(* IEC 61131-3 sources: daoli-st-library/DL_Device (part 22) *)

(* ---- FB_DL_FilterSwitchLevel.st ---- *)
(*
  FB_DL_FilterSwitchLevel  —  过滤器液位/料位联锁（fail-safe LOW + 再生切换闭锁） / Filter level interlock with fail-safe LOW and regeneration interlock
  分类 Category : DL_Device
  版本 Version  : 1.0.0
  来源 Source   : t2-2-lbp — 液位联锁族零检索深化
  溯源 Origin   : clean-room 实现，未复制任何源码行
  功能 Function : 1) 传感器原始信号归一口径与 FB_DL_LevelSwitchVib 对齐（不实例化，
                  防抖上游承载）：TRUE = 介质覆盖叉体（料位高于低位）；归一取反后
                  TRUE = 低料位，防抖 tGlitch 后出 bLowLevel；
                  2) fail-safe LOW 语义：bEnable = FALSE（传感器失效/退出）→ 强制判
                  低料位（安全侧请求切换，防干转）；
                  3) 再生切换闭锁：bRegenActive 期间 + 结束后 tBlockAfter 窗内，
                  bSwReq 强制 FALSE（TOF 承载闭锁窗，闭锁沿用当拍量）；
                  4) 双表冗余可选：bRedundEn 且双表不一致持续 tDisTo → 故障级 03FE
                  独立锁存，失效安全侧强制判低。
  边界 Boundary : ① 组态闸：tGlitch/tDisTo/tBlockAfter 任一 <= 0 → 03FF 锁存；
                  ② 闭锁窗 TOF 无条件周期刷新（R7）；切换闭锁判据全当拍量；
                  ③ Device 段 0003 故障带收口：03FE/03FF 两格（分段理由见 InverterPdiPoll ②）；
                  ④ 无 GVL 依赖：纯引脚输入输出，无外部变量引用，无物理 IO 地址。
  依赖 Depends  : 与 FB_DL_LevelSwitchVib 归一口径语义对齐（不实例化）；Standard.library（TON / TOF / R_TRIG）
  码表 Error codes（Device 段 0003，窗口 041F~0421 / 故障 03FE~03FF）:
    16#0003_03FE 故障级：双表冗余失决（不一致持续 tDisTo），锁存至 bReset
    16#0003_03FF 故障级：组态非法（任一窗口域非法），锁存至 bReset
    16#0003_041F 信息级：低料位切换请求沿（bSwReq 首次 TRUE）
    16#0003_0420 信息级：再生闭锁激活（bRegenActive 期间请求被闭锁）
    16#0003_0421 信息级：冗余判定恢复正常沿（失决解除）
  修订历史 Revision :
    2026-11-19  v1.0.0  R41 首版（批次 4 · 序号 2）
*)

FUNCTION_BLOCK FB_DL_FilterSwitchLevel
VAR_INPUT
    bLvlRaw1     : BOOL := FALSE;     // 主表原始信号，TRUE = 介质覆盖叉体 [-] / Primary raw switch, TRUE = covered
    bLvlRaw2     : BOOL := TRUE;      // 备表原始信号（冗余可选），默认与主表一致口径 [-] / Secondary raw switch
    bRedundEn    : BOOL := FALSE;     // 双表冗余使能 [-] / Redundancy enable
    bRegenActive : BOOL := FALSE;     // 再生进行中 [-] / Regeneration active
    tGlitch      : TIME := T#500MS;   // 低料位确认防抖 [ms]，域 > 0 / Low-level debounce
    tDisTo       : TIME := T#2S;      // 冗余失决窗 [ms]，域 > 0 / Redundancy disagreement window
    tBlockAfter  : TIME := T#5S;      // 再生结束后闭锁延时 [ms]，域 > 0 / Post-regen interlock delay
    bEnable      : BOOL := TRUE;      // 传感器处理使能，FALSE = 失效安全侧 [-] / Sensor enable, FALSE = fail-safe
    bReset       : BOOL := FALSE;     // 复位，上升沿清故障锁存 / Reset edge clears fault latch
END_VAR
VAR_OUTPUT
    bLowLevel    : BOOL;              // 归一低料位判定（fail-safe 口径）[-] / Normalized low-level verdict
    bSwReq       : BOOL;              // 再生切换请求（闭锁窗内强制 FALSE）[-] / Switch request, forced off in interlock
    bBlock       : BOOL;              // 闭锁窗激活标志 [-] / Interlock active flag
    bError       : BOOL;              // 故障锁存标志 / Fault latch flag
    nErrId       : UDINT;             // 事件码，0 = 无事件 / Event code
END_VAR
VAR
    tonLowDeb    : TON;               // 低料位防抖定时器，无条件周期刷新 / Low-level debounce timer
    tonDisTo     : TON;               // 冗余失决定时器（专用超时命名），无条件刷新 / Disagreement timer
    tofBlock     : TOF;               // 再生闭锁窗（TOF 承载再生后延时），无条件刷新 / Post-regen interlock timer
    rtReset      : R_TRIG;            // 复位沿实例，无条件刷新 / Reset edge instance
    _bLowNorm    : BOOL;              // 归一低料位当拍量（取反口径）/ Normalized low-level flag
    _bDisagree   : BOOL;              // 双表不一致当拍量 [-] / Disagreement current-scan flag
    _bDisLat     : BOOL;              // 失决锁存位（锁存量）/ Disagreement latch bit
    _bCfgBad     : BOOL;              // 组态锁存位（锁存量）/ Config-fault latch bit
    _uFault      : UDINT;             // 故障码锁存（锁存量）/ Latched fault code
    _uInfo       : UDINT;             // 信息码，每拍重算 / Transient info code
    _bSwReqPrev  : BOOL;              // 上拍请求镜像（请求沿判据）/ Previous request mirror
    _bBlockPrev  : BOOL;              // 上拍闭锁镜像（闭锁沿判据）/ Previous block mirror
    _bDisOkPrev  : BOOL;              // 上拍一致镜像（恢复沿判据）/ Previous agreement mirror
END_VAR

(* —— 段 0：定时器与沿实例无条件周期刷新（禁置于 IF/CASE 内） —— *)
_bLowNorm := NOT bLvlRaw1;                    // 归一取反：TRUE = 低料位（当拍量）
_bDisagree := bRedundEn AND (bLvlRaw1 <> bLvlRaw2);   // 双表不一致（当拍量）
rtReset(CLK := bReset);                       // 复位沿（每拍必调）
tonLowDeb(IN := _bLowNorm AND (NOT _bDisLat), PT := tGlitch);   // 低料位防抖（每拍必调）
tonDisTo(IN := _bDisagree, PT := tDisTo);     // 失决窗（每拍必调）
tofBlock(IN := bRegenActive, PT := tBlockAfter);  // 闭锁窗（再生期间 + 再生后延时，每拍必调）

(* —— 段 1：单拍量预清零（锁存量 _uFault/_bDisLat/_bCfgBad 不入清单，禁同拍抹除） —— *)
_uInfo := 16#0000_0000;             // 信息码每拍重算
nErrId := 16#0000_0000;             // 事件码缺省无事件

(* —— 段 2：复位沿 + 组态域闸（当拍量判据） —— *)
IF rtReset.Q THEN                   // rtReset.Q = 当拍量
    _bDisLat := FALSE;              // 清失决锁存位
    _bCfgBad := FALSE;              // 清组态锁存位
    _uFault := 16#0000_0000;        // 清故障锁存码
END_IF
IF (TIME_TO_DINT(tGlitch) <= 0) OR (TIME_TO_DINT(tDisTo) <= 0) OR (TIME_TO_DINT(tBlockAfter) <= 0) THEN
    _uFault := 16#0003_03FF;        // 故障级：组态非法
    _bCfgBad := TRUE;
END_IF

(* —— 段 3：冗余失决独立锁存与恢复（R190：失决归因唯一） —— *)
IF tonDisTo.Q AND (NOT _bDisLat) THEN
    _uFault := 16#0003_03FE;        // 故障级：双表失决锁存
    _bDisLat := TRUE;
END_IF
(* 解除式逐 BOOL 标注（R240）：rtReset.Q = 当拍量；NOT _bDisagree = 当拍量；
   均不含锁存量（_bDisLat），解除边真实可达。 *)
IF rtReset.Q AND (NOT _bDisagree) AND (NOT _bCfgBad) THEN
    _bDisLat := FALSE;              // 清失决锁存位（锁存量，仅此当拍量解除沿可清）
    _uFault := 16#0000_0000;        // 清故障锁存码（锁存量，同上唯一解除路径）
END_IF
IF (NOT _bDisagree) AND _bDisOkPrev AND bRedundEn AND (NOT _bDisLat) THEN
    _uInfo := 16#0003_0421;         // 信息级：冗余判定恢复沿
END_IF

(* —— 段 4：fail-safe LOW 归一出口（失效/失决/组态坏 → 强制判低，安全侧） —— *)
IF (NOT bEnable) OR _bDisLat OR _bCfgBad THEN
    bLowLevel := TRUE;              // 安全侧强制判低（防干转，头注释②）
ELSE
    bLowLevel := tonLowDeb.Q;       // 防抖后低料位判定
END_IF

(* —— 段 5：再生切换闭锁（闭锁判据全当拍量；TOF 电平承载再生后窗） —— *)
bBlock := bRegenActive OR tofBlock.Q;   // 闭锁窗激活（再生中或再生后延时内）
bSwReq := bLowLevel AND (NOT bBlock);   // 切换请求（闭锁窗内强制 FALSE）
IF bBlock AND (NOT _bBlockPrev) THEN
    _uInfo := 16#0003_0420;         // 信息级：再生闭锁激活
END_IF
IF bSwReq AND (NOT _bSwReqPrev) THEN
    _uInfo := 16#0003_041F;         // 信息级：切换请求沿（覆盖闭锁沿，请求优先报告）
END_IF

(* —— 段 6：出口单点映射（锁存码回放，禁同拍抹除） —— *)
IF _bDisLat OR _bCfgBad THEN
    nErrId := _uFault;              // 故障锁存码回放
ELSE
    nErrId := _uInfo;               // 信息码
END_IF
bError := _bDisLat OR _bCfgBad;     // 故障标志与锁存位同源
_bSwReqPrev := bSwReq;              // 请求沿判据快照
_bBlockPrev := bBlock;              // 闭锁沿判据快照
_bDisOkPrev := NOT _bDisagree;      // 一致镜像快照

END_FUNCTION_BLOCK

(* ---- FB_DL_FlowSwitchResponseCheck.st ---- *)
(*==============================================================================
 * 组件名称 (Component)  : FB_DL_FlowSwitchResponseCheck
 * 所属子库 (Sublibrary) : DL_Device
 * 当前版本 (Version)    : 1.0.0
 * 兼容性   (Platform)   : CODESYS 3.5+ / TwinCAT 3 / 汇川 InoProShop / 施耐德 Machine Expert
 *                         仅依赖 Standard.library（TON / R_TRIG），零厂商私有库
 * 功能描述 (Function)   : 流量开关**自身响应**校核（命令-监视-判定三段式）。① 运行指令 bRunCmd
 *                         上升沿起，tRespWin 内应出现流量开关 bFlowSw 上升沿；未出现 →
 *                         eCause = eNoResponse（开关卡死 / 管路堵塞 / 接线断）；② 指令撤销后
 *                         tDropWin 内流量信号未回落 → eCause = eStuckOn（开关粘连，常闭触点焊死）。
 *                         另输出实测响应时间 tRespMeasured（供趋势与开关劣化判断）。
 * 分工声明 (Scope)      : 本件**不判干转**（干转属主为 `FB_DL_PumpDryRunGuard` /
 *                         `FB_DL_PumpDryRunProtect`），也不判流量大小与累计量；本件只判「开关
 *                         是否按命令跟上、是否按命令放开」。干转保护需要泵曲线与最小流量阈值，
 *                         语义与本件正交，禁止互相替代。
 * 接口     (Interface)  : 输入 bRunCmd 泵/阀运行指令、bFlowSw 流量开关反馈、tRespWin 响应窗、
 *                         tDropWin 回落窗、bReset 复位；输出 bSwHealthy 开关健康位、tRespMeasured
 *                         实测响应时间（ET 锁存式）、eCause 归因、eState / bError / nErrId。
 * 边界     (Boundary)   : ① 组态闸：tRespWin <= T#0S 或 tDropWin <= T#0S → 故障锁存；
 *                         ② 响应时间测量用 **TON 的 ET 锁存**（流量沿那一拍读一次 ET 并锁存，
 *                         之后不再实时读 ET——锁存后实例继续计时会把测量值篡改，R38 范式）；
 *                         ③ TON 两枚 + R_TRIG 三枚段 0 无条件周期刷新，IN 由相位派生（R228A）；
 *                         ④ 故障相迁出唯一路径 = bReset 上升沿；⑤ 零全局耦合（无 GVL / 无物理地址）。
 * 解除式   (Release)    : bReset 上升沿 ∧ 组态合法 ∧ 当拍「指令与反馈同相」（bRunCmd 与 bFlowSw
 *                         同为真或同为假，即不处于任一异常窗，全为当拍量，R240 范式）。
 *                         自证可满足（终审两式 1）：两枚 TON 的 IN 挂相位，故障相内恒假 → Q 恒假；
 *                         现场消除卡死或粘连后指令与反馈自然同相，无恒假因子。
 * 码表     (Codes)      : 16#0003_0703 故障级：流量开关响应故障总码（组态非法 / 无响应 / 粘连 /
 *                         非法相位），锁存至 bReset 上升沿，归因由 eCause 承载（R190 单件单总码）；
 *                         16#0003_0482 信息级：响应正常（本次启动已在窗内测到响应沿）。
 *                         加码反证（R90）：响应正常时 tRespMeasured 已给出数值，但「本次启动已确认
 *                         响应」与「上一轮遗留的旧响应时间」在出口上无法区分（时间量会保持），
 *                         故立一码标记本轮已确认。
 *                         码段说明：Device 的 03xx 故障子带已占满（仅余 03C5~03C9 碎片孔洞，按
 *                         实战规则 13 禁回填），故本批新开 07xx 故障子带取 16#0003_0703；
 *                         信息级用 04xx 子带取 16#0003_0482（源码实扫为空）。分段理由即此。
 * 开源溯源 (Origin)     : 道莅自研 clean-room（参考命令-监视-判定三段式与参数域，
 *                         零代码行复制；t2-2-lbp 族）
 * 修订历史 (Revision)   : 2026-11-19  v1.0.0  R45 首版（批次 4 · 序号 17）
 *==============================================================================*)

TYPE E_DL_FsrState :
(
    eIdle     := 0,     // 待机（指令撤销且反馈已回落） / Idle, command off and feedback dropped
    eRespWait := 10,    // 响应窗内等流量信号 / Waiting for flow signal inside the response window
    eRun      := 20,    // 指令在效且流量已建立 / Command on and flow established
    eDropWait := 30,    // 回落窗内等流量信号消失 / Waiting for flow signal to drop inside the drop window
    eFault    := 90     // 故障锁存相 / Fault latched phase
);
END_TYPE

TYPE E_DL_FsrCause :
(
    eNone       := 0,   // 无故障成因 / No cause
    eCfgIllegal := 1,   // 组态非法 / Illegal configuration
    eNoResponse := 2,   // 无响应（窗内无流量沿） / No response inside the window
    eStuckOn    := 3,   // 粘连（撤销后不回落） / Stuck on, no drop after release
    ePhaseBad   := 4    // 非法相位兜底 / Illegal phase fallback
);
END_TYPE

FUNCTION_BLOCK FB_DL_FlowSwitchResponseCheck
VAR_INPUT
    bRunCmd    : BOOL := FALSE;          // 泵/阀运行指令（电平） [-] / Pump or valve run command level
    bFlowSw    : BOOL := FALSE;          // 流量开关反馈 [-] / Flow switch feedback
    tRespWin   : TIME := T#3S;           // 响应窗（指令起算），域 > T#0S [ms] / Response window, domain > T#0S [ms]
    tDropWin   : TIME := T#3S;           // 回落窗（撤令起算），域 > T#0S [ms] / Drop window, domain > T#0S [ms]
    bReset     : BOOL := FALSE;          // 复位命令，上升沿清故障 [-] / Reset command, rising edge clears fault
END_VAR
VAR_OUTPUT
    bSwHealthy   : BOOL;                 // 开关健康位（无故障且不在异常窗） [-] / Switch healthy flag
    tRespMeasured: TIME;                 // 实测响应时间（ET 锁存，锁存后不随实例计时变化） [ms] / Measured response time, latched ET [ms]
    eCause       : E_DL_FsrCause;        // 故障成因出口（R190 归因唯一） / Fault cause outlet
    eState       : E_DL_FsrState;        // 状态出口，段 6 单点映射 / State outlet
    bError       : BOOL;                 // 故障锁存标志 [-] / Fault latch flag
    nErrId       : UDINT;                // 事件码，0 = 无事件 / Event code, 0 = no event
END_VAR
VAR
    _eState      : E_DL_FsrState := E_DL_FsrState.eIdle;     // 内部相位（CASE 唯一写入目标） / Internal phase
    _eCause      : E_DL_FsrCause := E_DL_FsrCause.eNone;     // 故障成因锁存（锁存量） / Latched cause
    tonResp      : TON;                  // 响应窗计时，段 0 无条件调用 / Response window timer
    tonDrop      : TON;                  // 回落窗计时，段 0 无条件调用 / Drop window timer
    rtRun        : R_TRIG;               // 指令上升沿实例，段 0 无条件调用 / Command rising edge
    rtFlow       : R_TRIG;               // 流量上升沿实例，段 0 无条件调用 / Flow rising edge
    rtReset      : R_TRIG;               // 复位沿实例，段 0 无条件调用 / Reset edge
    _tRespLatch  : TIME;                 // 响应时间锁存槽（锁存量） [ms] / Response time latch, latched
    _bRespSeen   : BOOL;                 // 本轮已测到响应沿标记（锁存量） [-] / Response-seen flag for this run
    _bCfgBad     : BOOL;                 // 组态非法当拍量 [-] / Illegal configuration
    _bSamePhase  : BOOL;                 // 指令与反馈同相当拍量 [-] / Command and feedback in the same phase
    _bFault      : BOOL;                 // 故障锁存位（锁存量） / Latched fault bit
    _uFault      : UDINT;                // 故障码锁存（锁存量） / Latched fault code
    _uInfo       : UDINT;                // 信息码，每拍重算 / Info code, recomputed each scan
END_VAR

(* —— 段 0：当拍判据派生 + 定时器与沿实例无条件周期刷新 —— *)
_bCfgBad    := (tRespWin <= T#0S) OR (tDropWin <= T#0S);                            // 组态域闸 / Configuration gate
_bSamePhase := (bRunCmd AND bFlowSw) OR ((NOT bRunCmd) AND (NOT bFlowSw));           // 指令与反馈同相 / Command and feedback in the same phase
rtRun(CLK := bRunCmd);                                                              // 指令上升沿，每拍必调（R228A） / Command rising edge
rtFlow(CLK := bFlowSw);                                                             // 流量上升沿，每拍必调 / Flow rising edge
rtReset(CLK := bReset);                                                             // 复位沿，每拍必调 / Reset edge
tonResp(IN := (_eState = E_DL_FsrState.eRespWait), PT := tRespWin);                 // 响应窗计时（IN 由相位派生） / Response window timer
tonDrop(IN := (_eState = E_DL_FsrState.eDropWait), PT := tDropWin);                 // 回落窗计时 / Drop window timer

(* —— 段 1：单拍量预清零（锁存量不入清单，R107） —— *)
_uInfo       := 16#0000_0000;      // 信息码每拍重算 / Info recomputed every scan
bSwHealthy   := FALSE;             // 健康位每拍预清 / Healthy flag preset
tRespMeasured := _tRespLatch;      // 响应时间镜像（锁存量回放，不实时读 ET） / Response time mirror from the latch
nErrId       := 16#0000_0000;      // 事件码缺省无事件 / Event code default none
bError       := FALSE;             // 故障标志每拍预清，故障分支同拍置位（R45 配对） / Flag preset

(* —— 段 2：复位沿 + 组态域闸 —— *)
IF rtReset.Q THEN                                                        // 当拍复位沿 / current-scan reset edge
    _bFault := FALSE;                                                    // 清故障锁存位（锁存量） / Clear fault latch
    _uFault := 16#0000_0000;                                             // 清故障锁存码（锁存量） / Clear latched code
    _eCause := E_DL_FsrCause.eNone;                                      // 清成因（锁存量） / Clear latched cause
    IF _eState = E_DL_FsrState.eFault THEN
        _eState := E_DL_FsrState.eIdle;                                  // 故障相迁出唯一路径 / Sole exit from fault phase
    END_IF
END_IF
IF _bCfgBad THEN                                                         // 组态域闸 / Configuration gate
    _uFault := 16#0003_0703;                                             // 故障级：流量开关响应故障总码 / Fault-level: flow-switch fault code
    _bFault := TRUE;
    bError  := TRUE;                                                     // 故障标志同拍置位（R45 配对） / Error flag set same scan
    _eCause := E_DL_FsrCause.eCfgIllegal;                                // 归因：组态非法 / Cause: illegal configuration
END_IF

(* —— 段 3：响应时间测量（ET 只在流量沿那一拍读一次并锁存，R38 范式） —— *)
IF (NOT _bFault) AND (_eState = E_DL_FsrState.eRespWait) AND rtFlow.Q THEN
    _tRespLatch := tonResp.ET;                                           // 锁存响应时间（此后不再实时读 ET） / Latch ET once, never re-read live
    _bRespSeen := TRUE;                                                  // 本轮已确认响应 / Response confirmed for this run
    _uInfo := 16#0003_0482;                                              // 信息级：响应正常 / Info: response OK
END_IF

(* —— 段 4：无响应 / 粘连双判据（各用独立实例与独立归因，R190） —— *)
IF (NOT _bFault) AND tonResp.Q THEN                                      // 响应窗内无流量沿 → 无响应 / No flow edge inside the window
    _uFault := 16#0003_0703;
    _bFault := TRUE;
    bError  := TRUE;
    _eCause := E_DL_FsrCause.eNoResponse;                                // 归因：无响应 / Cause: no response
END_IF
IF (NOT _bFault) AND tonDrop.Q THEN                                      // 回落窗内流量未消失 → 粘连 / Flow did not drop inside the window
    _uFault := 16#0003_0703;
    _bFault := TRUE;
    bError  := TRUE;
    _eCause := E_DL_FsrCause.eStuckOn;                                   // 归因：粘连 / Cause: stuck on
END_IF

(* —— 段 5：故障解除式（R240 全当拍量） —— *)
IF rtReset.Q AND (NOT _bCfgBad) AND _bSamePhase THEN
    _bFault := FALSE;                                                    // 清故障锁存位（锁存量） / Clear fault latch
    _uFault := 16#0000_0000;                                             // 清故障锁存码（锁存量） / Clear latched code
    _eCause := E_DL_FsrCause.eNone;                                      // 清成因（锁存量） / Clear latched cause
END_IF

(* —— 段 5A：故障锁存相位迁移闸 —— *)
IF _bFault AND (_eState <> E_DL_FsrState.eFault) THEN
    _eState := E_DL_FsrState.eFault;                                     // 锁存即入故障相 / Latch enters fault phase
END_IF

(* —— 段 6：相位机（ENUM 全成员显式标签 + ELSE 兜底，R128） —— *)
CASE _eState OF

E_DL_FsrState.eIdle:
    IF rtRun.Q AND (NOT _bFault) THEN                                    // 出口 1：收到运行指令 / Run command received
        _bRespSeen := FALSE;                                             // 新一轮响应测量重新武装 / Re-arm response measurement
        _eState := E_DL_FsrState.eRespWait;
    ELSIF bFlowSw AND (NOT bRunCmd) THEN                                 // 出口 2：无令而流量已在（越序，交由回落链监视） / Flow on without command
        _eState := E_DL_FsrState.eDropWait;
    ELSIF _bFault THEN                                                   // 出口 3：故障锁存 / Fault latched
        _eState := E_DL_FsrState.eFault;
    END_IF

E_DL_FsrState.eRespWait:
    IF rtFlow.Q THEN                                                     // 出口 1：窗内出现流量沿 / Flow edge inside the window
        _eState := E_DL_FsrState.eRun;
    ELSIF NOT bRunCmd THEN                                               // 出口 2：指令撤销（前置消失，R98） / Command released
        _eState := E_DL_FsrState.eIdle;
    END_IF

E_DL_FsrState.eRun:
    IF NOT bRunCmd THEN                                                  // 出口 1：撤销指令，进回落窗 / Command released, enter drop window
        _eState := E_DL_FsrState.eDropWait;
    ELSIF NOT bFlowSw THEN                                               // 出口 2：运行中流量消失（前置消失，R98） / Flow lost while running
        _eState := E_DL_FsrState.eRespWait;
    END_IF

E_DL_FsrState.eDropWait:
    IF NOT bFlowSw THEN                                                  // 出口 1：流量已回落 / Flow dropped
        _eState := E_DL_FsrState.eIdle;
    ELSIF bRunCmd THEN                                                   // 出口 2：指令重新来（前置消失，R98） / Command came back
        _eState := E_DL_FsrState.eRespWait;
    END_IF

E_DL_FsrState.eFault:
    ;                                                                     // 故障相：仅段 5 复位沿可迁出 / Only the reset edge leaves this phase

ELSE
    _uFault := 16#0003_0703;                                             // 故障级：非法相位兜底（归并总码） / Illegal-phase fallback
    _bFault := TRUE;
    bError  := TRUE;
    _eCause := E_DL_FsrCause.ePhaseBad;                                  // 归因：非法相位 / Cause: illegal phase
    _eState := E_DL_FsrState.eFault;

END_CASE

(* —— 段 7：出口单点映射（名实同源；锁存码回放） —— *)
bSwHealthy := (NOT _bFault) AND _bSamePhase AND _bRespSeen;              // 健康 = 无故障 ∧ 同相 ∧ 本轮已确认响应 / Healthy verdict
IF _bFault THEN
    nErrId := _uFault;                                                   // 故障锁存码回放 / Replay latched fault code
ELSE
    nErrId := _uInfo;                                                    // 信息码 / Info code
END_IF
bError := _bFault;                                                       // 故障标志与锁存同源（名实双出口，R191） / Flag from latch
eState := _eState;                                                       // 状态出口 / State outlet
eCause := _eCause;                                                       // 成因出口 / Cause outlet

END_FUNCTION_BLOCK

(* ---- FB_DL_FoupDoorSeq.st ---- *)
// =====================================================================
// FB_DL_FoupDoorSeq.st
// FOUP 开合门与载具联锁顺控（解锁-开门-载具在位-再锁定确认窗）
// FOUP door interlock sequencing with relock confirm window
// 所属子库: DL_Device    版本: v1.0.0    兼容: CODESYS V3.5+ / TwinCAT 3 / 汇川 InoProShop
// 码位: 16#0003_03DE ~ 16#0003_03E2 (本件独占 5 槽, 勿复用)
// 溯源: 道莅 clean-room 防御性实现
//       来源组标签: semiconductor, door-interlock, sequencing, foup
// 枚举属主: E_DL_FoupDoorState —— 本文件为全库唯一属主, 其他件只引用不重声明
// 修改记录: R30 初版 (ROUND_PLAN_R30 序 2)
// =====================================================================
// ---------------------------------------------------------------------
// 枚举定义: E_DL_FoupDoorState (全库唯一属主, 其他件只引用不重声明)
// ---------------------------------------------------------------------
TYPE E_DL_FoupDoorState :
(
    eIdle,          // 空闲（门锁闭等待）/ Idle, locked
    eUnlocking,     // 解锁保持中 / Unlocking
    eDoorOpen,      // 门已开等待传输 / Door open
    eTransfer,      // 载具传输中 / Transfer in progress
    eRelocking,     // 再锁定确认窗 / Relocking confirm window
    eFault          // 故障锁存 / Fault latched
);
END_TYPE

FUNCTION_BLOCK FB_DL_FoupDoorSeq
VAR_INPUT
    bEnable         : BOOL  := FALSE;   // 使能 / Enable
    bDoorClosed     : BOOL  := FALSE;   // 门磁关到位反馈 / Door closed feedback
    bDoorOpen       : BOOL  := FALSE;   // 门磁开到位反馈 / Door open feedback
    bCarrierPresent : BOOL  := FALSE;   // 载具在位检测 / Carrier present detection
    bUnlockCmd      : BOOL  := FALSE;   // 解锁命令 / Unlock command
    bLockCmd        : BOOL  := FALSE;   // 锁定命令 / Lock command
    bVacuumOk       : BOOL  := FALSE;   // 真空解锁条件就绪 / Vacuum release ready
    tUnlockHold     : TIME  := T#3S;    // 解锁保持超时窗 T#100MS~T#60S / Unlock hold timeout window [s]
    tRelockWin      : TIME  := T#5S;    // 再锁定确认窗 T#100MS~T#60S / Relock confirm window [s]
    bReset          : BOOL  := FALSE;   // 故障复位命令 / Fault reset command
END_VAR
VAR_OUTPUT
    bUnlockOut      : BOOL := FALSE;    // 解锁输出, 安全侧为假 / Unlock output, safe side FALSE
    bLockOut        : BOOL := FALSE;    // 锁定输出 / Lock output
    eState          : E_DL_FoupDoorState := E_DL_FoupDoorState.eIdle;  // 顺控状态 / Sequence state
    bTransferPermit : BOOL := FALSE;    // 载具传输允许 / Transfer permit
    eErr            : UDINT := 16#0003_03DE;  // 错误码 / Error code
END_VAR
VAR
    eErrLatch       : UDINT := 16#0003_03DE;  // 故障锁存码回放 / Latched fault code replay
    bDoorConflict   : BOOL := FALSE;    // 门磁双反馈矛盾 / Door feedback conflict
    rtrReset        : R_TRIG;           // 复位上升沿检测, 每拍无条件刷新 / Reset edge, refreshed every cycle
    tonUnlock       : TON;              // 解锁保持超时定时器, 每拍无条件刷新 / Unlock hold timer, refreshed every cycle
    tonRelock       : TON;              // 再锁定确认窗定时器, 每拍无条件刷新 / Relock window timer, refreshed every cycle
END_VAR

// ---------------------------------------------------------------------
// 代码位表（本件独占, 勿复用）:
//   16#0003_03DE 信息 顺控正常（空闲或顺控执行中）
//   16#0003_03DF 故障 解锁保持超时（解锁输出有效而门未开超时）, 解除式 = bReset 上升沿 且 门磁回到关到位 且 无矛盾反馈
//   16#0003_03E0 故障 再锁定确认窗超时（窗内门磁未回关到位）, 解除式同 03DF
//   16#0003_03E1 故障 门磁双反馈矛盾（关到位与开到位同时有效）, 解除式同 03DF
//   16#0003_03E2 故障 非法状态兜底（状态机 ELSE 拦截）, 解除式同 03DF
// ---------------------------------------------------------------------

// ---- 门磁矛盾判（最高优先级拦截）/ Door feedback conflict: highest priority ----
bDoorConflict := bDoorClosed AND bDoorOpen;     // 双反馈同有效 = 组态或接线矛盾 / Both active = conflict
IF bDoorConflict THEN
    eState    := E_DL_FoupDoorState.eFault;     // 任意相直接落故障 / Fall to fault from any phase
    eErrLatch := 16#0003_03E1;                  // 锁存矛盾码 / Latch conflict code
END_IF

// ---- 非故障相下使能撤销 → 回空闲（安全侧）/ Disable in non-fault phase returns to idle ----
IF (NOT bEnable) AND (eState <> E_DL_FoupDoorState.eFault) THEN
    eState := E_DL_FoupDoorState.eIdle;         // 退回空闲 / Return to idle
END_IF

// ---- 定时器与边沿实例无条件周期刷新（调用本身不进任何 IF 分支）/ Unconditional timer and edge refresh ----
tonUnlock(IN := (eState = E_DL_FoupDoorState.eUnlocking) AND (NOT bDoorOpen),
          PT := tUnlockHold);                   // 解锁保持计时 / Unlock hold timing
tonRelock(IN := (eState = E_DL_FoupDoorState.eRelocking) AND (NOT bDoorClosed),
          PT := tRelockWin);                    // 再锁定确认窗计时 / Relock window timing
rtrReset(CLK := bReset);                        // 复位沿检测 / Reset edge detection

// ---- 默认输出（安全侧全 0, 各相按需覆盖）/ Default outputs (safe side) ----
bUnlockOut      := FALSE;   // 解锁输出缺省断开 / Unlock default off
bLockOut        := FALSE;   // 锁定输出缺省断开 / Lock default off
bTransferPermit := FALSE;   // 传输允许缺省禁止 / Permit default denied

// ---- 状态机 / State machine ----
IF eState = E_DL_FoupDoorState.eFault THEN
    // 故障相: 输出全 0, 锁存码回放 / Fault phase: outputs all off, latch replay
    eErr := eErrLatch;
    // 解除式: bReset 上升沿 且 门磁回到关到位 且 无矛盾反馈 / Release: reset edge AND closed AND no conflict
    IF rtrReset.Q AND bDoorClosed AND (NOT bDoorOpen) AND (NOT bDoorConflict) THEN
        eState    := E_DL_FoupDoorState.eIdle;  // 解除故障回空闲 / Release to idle
        eErrLatch := 16#0003_03DE;              // 清锁存码 / Clear latch code
    END_IF
ELSE
    CASE eState OF
        E_DL_FoupDoorState.eIdle:       // 空闲: 门锁闭等待解锁命令 / Idle: locked, wait unlock
            bLockOut := bDoorClosed;    // 锁定输出随关到位反馈 / Lock output follows closed feedback
            IF bUnlockCmd AND bVacuumOk AND (NOT bDoorConflict) THEN
                eState := E_DL_FoupDoorState.eUnlocking;    // 拍 N 进入解锁相 / Enter unlocking
            END_IF
        E_DL_FoupDoorState.eUnlocking:  // 解锁保持: 输出有效等待门开 / Unlocking: output on, wait door open
            bUnlockOut := TRUE;         // 解锁输出有效 / Unlock output on
            // 本拍行为: 门开转开门相, 真空条件丢失回空闲, 超时落故障 / Open to door phase, vacuum loss to idle, timeout to fault
            IF bDoorOpen AND (NOT bDoorConflict) THEN
                eState := E_DL_FoupDoorState.eDoorOpen;     // 拍 N+1 转开门相 / To door-open phase
            ELSIF NOT bVacuumOk THEN
                eState := E_DL_FoupDoorState.eIdle;         // 真空条件丢失中止解锁 / Vacuum lost, abort unlock
            ELSIF tonUnlock.Q THEN
                eState    := E_DL_FoupDoorState.eFault;     // 解锁有效但门未开超时 / Unlock valid but not open in time
                eErrLatch := 16#0003_03DF;                  // 锁存超时码 / Latch timeout code
            END_IF
        E_DL_FoupDoorState.eDoorOpen:   // 门已开: 允许传输, 等载具在位或锁定命令 / Door open: permit, wait carrier or lock cmd
            bUnlockOut      := TRUE;    // 开门期间保持解锁 / Hold unlock while open
            bTransferPermit := TRUE;    // 允许载具传输 / Permit transfer
            IF bCarrierPresent THEN
                eState := E_DL_FoupDoorState.eTransfer;     // 载具在位转传输相 / Carrier present, to transfer
            ELSIF bLockCmd AND (NOT bDoorConflict) THEN
                eState := E_DL_FoupDoorState.eRelocking;    // 直接收到锁定命令转确认窗 / Lock cmd, to relocking
            END_IF
        E_DL_FoupDoorState.eTransfer:   // 载具传输中: 保持允许, 等锁定命令 / Transfer: permit held, wait lock cmd
            bUnlockOut      := TRUE;    // 传输期间保持解锁 / Hold unlock during transfer
            bTransferPermit := TRUE;    // 保持传输允许 / Hold transfer permit
            IF bLockCmd AND (NOT bDoorConflict) THEN
                eState := E_DL_FoupDoorState.eRelocking;    // 收到锁定命令转确认窗 / Lock cmd, to relocking
            END_IF
        E_DL_FoupDoorState.eRelocking:  // 再锁定确认窗: 门磁必须回关到位 / Relocking: door must return closed
            bLockOut := TRUE;           // 锁定输出有效 / Lock output on
            // 本拍行为: 门关到位转空闲, 窗超时落故障 / Closed to idle, window timeout to fault
            IF bDoorClosed AND (NOT bDoorConflict) THEN
                eState := E_DL_FoupDoorState.eIdle;     // 再锁定完成回空闲 / Relock done, to idle
            ELSIF tonRelock.Q THEN
                eState    := E_DL_FoupDoorState.eFault; // 确认窗内门磁未回关到位 / Door not closed in window
                eErrLatch := 16#0003_03E0;              // 锁存确认窗超时码 / Latch window timeout code
            END_IF
        ELSE                                    // 非法状态兜底拦截 / Illegal state fallback
            eState    := E_DL_FoupDoorState.eFault;     // 落故障相 / Fall to fault
            eErrLatch := 16#0003_03E2;                  // 锁存兜底码 / Latch fallback code
        END_CASE
    // 本拍错误码: 刚落故障则回放锁存码, 否则正常码 / Error code of this cycle
    IF eState = E_DL_FoupDoorState.eFault THEN
        eErr := eErrLatch;          // 回放锁存码 / Replay latch code
    ELSE
        eErr := 16#0003_03DE;       // 顺控正常 / Sequence normal
    END_IF
END_IF

END_FUNCTION_BLOCK

(* ---- FB_DL_FoupPurgeN2Flow.st ---- *)
(*
  FB_DL_FoupPurgeN2Flow  —  FOUP 氮气吹扫流量与露点监视（建立窗口 / 分级露点告警 / 注入脉冲流量计）/ FOUP N2 purge flow and dew-point supervision
  分类 Category : DL_Device
  码位 Code     : 16#03_2_0F
  版本 Version  : 1.0.0
  来源 Source   : t2-1-lgf-measurement — IEC 61131-3 标准语义的道莅防御性实现
  溯源 Origin   : LGF 测量类文档公开语义借鉴（流量带判据、露点分级），clean-room 实现，未复制源码行
  功能 Function : 1) 注入 FB_DL_PulseFlowMeter 实例（VAR_IN_OUT，只读其流量/总量/故障输出，**本件不调用其实例体**），
                     取瞬时流量与 K 系数参与判据；
                  2) 吹扫起始（bPurgeStart 上升沿）后在 tPurgeEstablish 内流量须进入 fFlowSetLpm ± fFlowTolPct% 带，
                     否则置 bEstablishTimeout（故障级 021F）；
                  3) 露点按两级判据告警：越 fDewPointMaxC 为「越限」（023F），越 fDewSevereC 为「严重越限」（024F），
                     两码独立、独立出口（R190 归因唯一）；
                  4) 露点信号质量坏或缺失时**不当作合格**：置 022F 且 bPurgeOk := FALSE（安全侧，绝不静默放行）。
  边界 Boundary : ① fFlowSetLpm <= 0 判组态错 020F（偏差百分比的分母，R45 防除零）；
                     注入流量计 fKFactor = 0 判组态错 020F 且不投运（K 系数未标定，流量读数无物理意义）；
                     露点两级门限倒置（fDewSevereC <= fDewPointMaxC）同判组态错；
                  ② 偏差百分比对 ABS 结果限幅 DL_DEV_CLAMP_PCT，防极端读数导致 REAL 溢出与 HMI 显示异常；
                  ③ bPurgeOk 的成立条件 = 建立成功 AND 流量在带 AND 露点未越限 AND 露点信号有效 AND 无故障；
                  ④ 解除式自证：_bFault 清除 = rtReset.Q（引脚可满足）；021F 另可由「流量重新入带且持续
                     tEstablishRetry」按码专清（R188 可达清除边）；023F/024F 可由露点回落按码专清；
                  ⑤ bDewPointAlarm / bDewSevereAlarm 为保持型告警位（不随单拍读数抖动），只由复位沿或回落清除。
  依赖 Depends  : FB_DL_PulseFlowMeter（DL_Device 既有件，×1 以 VAR_IN_OUT 注入）；
                  仅 Standard.library（TON / R_TRIG / ABS / MIN / MAX）
  同拍双窗配比  : tPurgeEstablish（建立窗口）与 tDewDb（露点去抖窗）不同源；配比约束
                  tDewDb <= tPurgeEstablish，保证建立窗口内露点结论至少更新一次（R100）

  码表 Error codes（本件格 03_2_0F，子码步进 +0x10）:
    16#0003_020F 故障级：组态非法（流量设定 <= 0 / K 系数 = 0 / 容差 <= 0 / 露点门限倒置 / 时间参数 <= 0）
    16#0003_021F 故障级：吹扫建立超时（tPurgeEstablish 内流量未进入容许带）
    16#0003_022F 故障级：露点信号无效（质量坏或缺失，不当作合格）
    16#0003_023F 故障级：露点越限（超 fDewPointMaxC）
    16#0003_024F 故障级：露点严重越限（超 fDewSevereC）
    16#0003_025F 故障级：状态机落 ELSE 兜底（非法相位 ID）
    16#0003_010F 信息级：吹扫建立成功，流量已入带（不置 bError）
    16#0003_011F 信息级：流量偏差瞬时越带但未超建立窗口（不置 bError）

  修订历史 Revision :
    2026-11-18  v1.0.0  R37 首版
*)

TYPE E_DL_N2PurgeState :
(
    eIdle      := 0,   // 空闲：未吹扫 / Idle, purge not started
    eEstablish := 10,  // 建立中：等流量进入容许带 / Establishing, waiting for the flow band
    ePurged    := 20,  // 吹扫中：流量与露点均在限内 / Purging, flow and dew point inside the limits
    eTimeout   := 30,  // 超时：建立窗口耗尽，等待复位 / Timed out, waiting for a reset
    eFault     := 90   // 故障：组态或信号故障锁定 / Fault, a latched configuration or signal fault
);
END_TYPE

FUNCTION_BLOCK FB_DL_FoupPurgeN2Flow
VAR_INPUT
    bEnable        : BOOL := FALSE;             // 总使能，FALSE 时 bPurgeOk 恒假 / Master enable, low level forces bPurgeOk FALSE
    bReset         : BOOL := FALSE;             // 复位，上升沿清故障与告警锁存 / Reset, clears the fault and alarm latches
    bPurgeStart    : BOOL := FALSE;             // 吹扫起始触发（上升沿受理）/ Purge start trigger, rising edge
    fFlowSetLpm    : REAL := 20.0;              // 吹扫流量设定 [L/min]，域 > 0 / Purge flow setpoint [L/min]
    fFlowTolPct    : REAL := 10.0;              // 流量容许带 [%]，域 > 0 / Flow tolerance band [%]
    fDewPointMaxC  : REAL := -40.0;             // 露点越限门限 [°C]，域 < fDewSevereC / Dew point limit [degC]
    fDewSevereC    : REAL := -20.0;             // 露点严重越限门限 [°C]，须 > fDewPointMaxC / Severe dew point limit [degC]
    fDewPointC     : REAL := -60.0;             // 露点实测值 [°C] / Measured dew point [degC]
    bDewQualityOk  : BOOL := TRUE;              // 露点信号质量（FALSE = 坏或缺失）/ Dew point signal quality, FALSE means bad
    tPurgeEstablish : TIME := T#10S;            // 吹扫建立窗口 [ms]，域 > 0 / Purge establishment window [ms]
    tEstablishRetry : TIME := T#30S;            // 入带持续窗（021F 按码专清用）[ms]，域 > 0 / In-band dwell for the code-specific clear
    tDewDb         : TIME := T#2S;              // 露点告警去抖窗 [ms]，域 > 0 / Dew point debounce [ms]
END_VAR
VAR_OUTPUT
    bPurgeOk       : BOOL;                      // 吹扫合格（建立成功且流量/露点均在限内）/ Purge acceptable
    bEstablishTimeout : BOOL;                   // 建立超时（保持型）/ Establishment timeout, held
    bDewPointAlarm : BOOL;                      // 露点越限告警（保持型）/ Dew point alarm, held
    bDewSevereAlarm : BOOL;                     // 露点严重越限告警（保持型）/ Severe dew point alarm, held
    fFlowDeviationPct : REAL;                   // 流量偏差 [%]，已限幅 / Flow deviation [%], clamped
    fFlowActualLpm : REAL;                      // 实测流量 [L/min] / Measured flow [L/min]
    bValid         : BOOL;                      // 判据可用标志 / Criteria usable
    bError         : BOOL;                      // 故障标志，派生自锁存 / Fault flag derived from the latch
    nErrId         : UDINT;                     // 事件码，0 = 无事件 / Event code, 0 = no event
    eStateOut      : E_DL_N2PurgeState;         // 状态出口，段尾单点映射 / State outlet, mapped at the tail
END_VAR
VAR_IN_OUT
    fbFlowMeter : FB_DL_PulseFlowMeter;         // 注入的脉冲流量计实例（只读输出，本件不调用其实例体）/ Injected pulse flow meter, read only
END_VAR
VAR
    tonEstablish : TON;                         // 建立窗口计时，每拍无条件调用 / Establishment window, called unconditionally
    tonInBand    : TON;                         // 入带持续计时，每拍无条件调用 / In-band dwell timer, called unconditionally
    tonDew       : TON;                         // 露点去抖计时，每拍无条件调用 / Dew point debounce, called unconditionally
    tonHeart     : TON;                         // 周期心跳窗，自复位 / Periodic heartbeat window, self-resetting
    rtReset      : R_TRIG;                      // 复位上升沿 / Reset rising edge
    rtStart      : R_TRIG;                      // 吹扫起始上升沿 / Purge start rising edge
    _eState      : E_DL_N2PurgeState := E_DL_N2PurgeState.eIdle;  // 内部相位（CASE 唯一写入目标）/ Internal phase
    _uFault      : UDINT;                       // 故障码锁存 / Latched fault code
    _uInfo       : UDINT;                       // 信息码，每拍重算 / Information code, recomputed per scan
    _bFault      : BOOL;                        // 故障锁存位 / Latched fault bit
    _bCfgBad     : BOOL;                        // 组态非法聚合 / Configuration invalid aggregate
    _bInBand     : BOOL;                        // 流量在容许带 / Flow inside the tolerance band
    _bEstTimeout : BOOL;                        // 建立超时保持量 / Held establishment-timeout value
    _bDewAlarm   : BOOL;                        // 露点越限保持量 / Held dew point alarm
    _bDewSevere  : BOOL;                        // 露点严重越限保持量 / Held severe dew point alarm
    _bDewBad     : BOOL;                        // 露点信号无效 / Dew point signal unusable
    _bEstBreak   : BOOL := TRUE;                // 建立窗口断输入一拍 / One-scan establishment break
    _bInBandBrk  : BOOL := TRUE;                // 入带计时断输入一拍 / One-scan in-band break
    _bDewBrk     : BOOL := TRUE;                // 露点去抖断输入一拍 / One-scan dew break
    _bHeartBrk   : BOOL := TRUE;                // 心跳窗断输入一拍 / One-scan heartbeat break
    _fDevRaw     : REAL;                        // 未限幅偏差 [%] / Unclamped deviation [%]
    _fKFactor    : REAL;                        // 注入流量计 K 系数 [pulses/L] / Injected K-factor [pulses/L]
END_VAR
VAR CONSTANT
    DL_DEV_CLAMP_PCT : REAL := 1000.0;   // 偏差绝对值限幅 [%] / Deviation magnitude clamp [%]
    DL_DEW_LIM_C     : REAL := 200.0;    // 露点有限性上限 [°C] / Dew point magnitude ceiling [degC]
    DL_FLOW_LIM_LPM  : REAL := 100000.0; // 流量有限性上限 [L/min] / Flow magnitude ceiling [L/min]
    DL_HEART_WINDOW  : TIME := T#2S;     // 心跳观察窗 [ms]，自复位节拍 / Heartbeat window, self-resetting
END_VAR

(* —— 段 0：定时器与边缘检测无条件周期刷新（R182：调用语句不得置于 IF / CASE 内） —— *)
rtReset(CLK := bReset);                                          // 复位上升沿，每拍必调
rtStart(CLK := bPurgeStart);                                     // 吹扫起始上升沿，每拍必调
tonHeart(IN := (NOT tonHeart.Q) AND (NOT _bHeartBrk), PT := DL_HEART_WINDOW);  // 心跳窗自复位
_bHeartBrk := FALSE;                                             // 断输入拍在调用后自清
tonEstablish(IN := (_eState = E_DL_N2PurgeState.eEstablish) AND (NOT _bEstBreak), PT := tPurgeEstablish);  // 建立窗口
_bEstBreak := FALSE;                                             // 断输入拍在调用后自清
tonInBand(IN := _bInBand AND (NOT _bInBandBrk), PT := tEstablishRetry);   // 入带持续（表达式入参）
_bInBandBrk := FALSE;                                            // 断输入拍在调用后自清
tonDew(IN := _bDewBad AND (NOT _bDewBrk), PT := tDewDb);          // 露点信号无效去抖（表达式入参）
_bDewBrk := FALSE;                                               // 断输入拍在调用后自清

(* —— 段 1：单拍量预清零（告警保持量 / 锁存不入清单，R187①） —— *)
_uInfo      := 16#0000_0000;   // 信息码每拍重算
bError      := FALSE;          // 故障出口每拍重算，段 6 由锁存派生
bValid      := FALSE;          // 可用标志缺省 FALSE
bPurgeOk    := FALSE;          // 合格出口缺省 FALSE（安全侧）
_bCfgBad    := FALSE;          // 组态非法预清零
_bInBand    := FALSE;          // 在带判据预清零
_bDewBad    := FALSE;          // 露点信号无效预清零

(* —— 段 2：复位沿清锁存与告警保持量（R188 双路径） —— *)
IF rtReset.Q THEN
    _bFault     := FALSE;            // 复位沿清锁存位
    _uFault     := 16#0000_0000;     // 复位沿清锁存码
    _bEstTimeout := FALSE;           // 清建立超时保持量
    _bDewAlarm  := FALSE;            // 清露点越限告警
    _bDewSevere := FALSE;            // 清露点严重越限告警
END_IF
IF (_uFault = 16#0003_023F) AND (NOT _bDewAlarm) THEN
    _uFault := 16#0000_0000;         // 按码专清：露点回落至越限门限以下
    _bFault := FALSE;                // 锁存位同步清
END_IF
IF (_uFault = 16#0003_024F) AND (NOT _bDewSevere) THEN
    _uFault := 16#0000_0000;         // 按码专清：露点回落至严重门限以下
    _bFault := FALSE;                // 锁存位同步清
END_IF

(* —— 段 3：组态域闸（覆盖全部参与换算的引脚与注入件参数，R151） —— *)
_fKFactor := fbFlowMeter.fKFactor;                              // 读注入件 K 系数 [pulses/L]
IF (fFlowSetLpm <> fFlowSetLpm) OR (fFlowSetLpm <= 0.0) OR (fFlowSetLpm > DL_FLOW_LIM_LPM) THEN
    _bCfgBad := TRUE;                                           // 流量设定非法（偏差分母，R45 防除零）
END_IF
IF (_fKFactor <> _fKFactor) OR (_fKFactor <= 0.0) THEN
    _bCfgBad := TRUE;                                           // K 系数未组态/非有限：流量读数无物理意义，不投运
END_IF
IF (fFlowTolPct <> fFlowTolPct) OR (fFlowTolPct <= 0.0) THEN
    _bCfgBad := TRUE;                                           // 容差带非法（为 0 等于永不合格）
END_IF
IF (fDewPointMaxC <> fDewPointMaxC) OR (ABS(fDewPointMaxC) > DL_DEW_LIM_C) THEN
    _bCfgBad := TRUE;                                           // 露点越限门限非法
END_IF
IF (fDewSevereC <> fDewSevereC) OR (fDewSevereC <= fDewPointMaxC) THEN
    _bCfgBad := TRUE;                                           // 严重门限倒置（须严格大于越限门限）
END_IF
IF (TIME_TO_DINT(tPurgeEstablish) <= 0) OR (TIME_TO_DINT(tEstablishRetry) <= 0) OR
   (TIME_TO_DINT(tDewDb) <= 0) THEN
    _bCfgBad := TRUE;                                           // 三个时间参数均须 > 0
END_IF
IF _bCfgBad THEN
    _uFault := 16#0003_020F;                                    // 故障级：组态非法
    _bFault := TRUE;                                            // 锁存位置位（复位沿可清）
    bError  := TRUE;                                            // 故障标志置位（R45 配对）
    _eState := E_DL_N2PurgeState.eFault;                        // 进故障相（不投运）
END_IF

(* —— 段 4：流量与露点判据（仅无组态错时计算） —— *)
IF NOT _bCfgBad THEN
    fFlowActualLpm := fbFlowMeter.fFlowRate;                    // 注入件瞬时流量镜像 [L/min]
    IF (fFlowActualLpm <> fFlowActualLpm) OR (ABS(fFlowActualLpm) > DL_FLOW_LIM_LPM) THEN
        _bCfgBad := TRUE;                                       // 流量非有限：本拍判据不可信
        _uFault := 16#0003_020F;                                // 故障级：输入异常归入组态/输入异常码
        _bFault := TRUE;                                        // 锁存
        bError  := TRUE;                                        // 故障标志置位（R45 配对）
        _eState := E_DL_N2PurgeState.eFault;                    // 进故障相
    ELSE
        _fDevRaw := (fFlowActualLpm - fFlowSetLpm) / fFlowSetLpm * 100.0;   // 偏差 [%]（分母已证 > 0）
        fFlowDeviationPct := _fDevRaw;                          // 出口初值
        IF fFlowDeviationPct > DL_DEV_CLAMP_PCT THEN
            fFlowDeviationPct := DL_DEV_CLAMP_PCT;              // 上行限幅（防溢出与显示异常）
        END_IF
        IF fFlowDeviationPct < -DL_DEV_CLAMP_PCT THEN
            fFlowDeviationPct := -DL_DEV_CLAMP_PCT;             // 下行限幅
        END_IF
        _bInBand := (ABS(_fDevRaw) <= fFlowTolPct);             // 在带判据（用未限幅偏差判，避免限幅掩盖超差）
        IF NOT _bInBand THEN
            _uInfo := 16#0003_011F;                             // 信息级：瞬时越带（可能仍可建立）
        END_IF
    END_IF

    (* 4A 露点信号质量：坏则**不当作合格**（安全侧） *)
    IF (NOT bDewQualityOk) OR (fDewPointC <> fDewPointC) OR (ABS(fDewPointC) > DL_DEW_LIM_C) THEN
        _bDewBad := TRUE;                                       // 信号无效
        _uFault := 16#0003_022F;                                // 故障级：露点信号无效
        _bFault := TRUE;                                        // 锁存
        bError  := TRUE;                                        // 故障标志置位（R45 配对）
    END_IF

    (* 4B 露点分级判据：越限 / 严重越限两码独立，保持型告警位 *)
    IF (NOT _bDewBad) THEN
        IF fDewPointC > fDewSevereC THEN
            _bDewSevere := TRUE;                                // 严重越限保持量
            _bDewAlarm  := TRUE;                                // 严重越限同时满足越限（上位包含关系）
            _uFault := 16#0003_024F;                            // 故障级：露点严重越限
            _bFault := TRUE;                                    // 锁存
            bError  := TRUE;                                    // 故障标志置位（R45 配对）
        ELSIF fDewPointC > fDewPointMaxC THEN
            _bDewAlarm := TRUE;                                 // 越限保持量
            _uFault := 16#0003_023F;                            // 故障级：露点越限
            _bFault := TRUE;                                    // 锁存
            bError  := TRUE;                                    // 故障标志置位（R45 配对）
        ELSE
            IF fDewPointC <= (fDewPointMaxC - 1.0) THEN
                _bDewAlarm := FALSE;                            // 回落 1 °C 回差：越限告警释放
            END_IF
            IF fDewPointC <= (fDewSevereC - 1.0) THEN
                _bDewSevere := FALSE;                           // 回落 1 °C 回差：严重告警释放
            END_IF
        END_IF
    END_IF
END_IF

(* —— 段 5：相位机（只做迁移；出口在段 7） —— *)
CASE _eState OF

E_DL_N2PurgeState.eIdle:
    IF rtStart.Q AND bEnable AND (NOT _bFault) AND (NOT _bCfgBad) THEN
        _eState := E_DL_N2PurgeState.eEstablish;      // 起始触发：进建立相
        _bEstBreak := TRUE;                          // 建立窗口从零计时
        _bInBandBrk := TRUE;                         // 入带计时从零
    END_IF

E_DL_N2PurgeState.eEstablish:
    IF (NOT bEnable) OR _bFault THEN
        _eState := E_DL_N2PurgeState.eFault;         // 失能或故障：进故障相（bPurgeOk 已为假）
    ELSIF _bInBand THEN
        _eState := E_DL_N2PurgeState.ePurged;        // 流量入带（含持续窗满）：进吹扫相
        _uInfo := 16#0003_010F;                      // 信息级：吹扫建立成功
    ELSIF tonEstablish.Q THEN
        _bEstTimeout := TRUE;                        // 建立超时保持量
        _uFault := 16#0003_021F;                     // 故障级：建立超时
        _bFault := TRUE;                             // 锁存
        bError  := TRUE;                             // 故障标志置位（R45 配对）
        _eState := E_DL_N2PurgeState.eTimeout;       // 进超时相
    END_IF

E_DL_N2PurgeState.ePurged:
    IF (NOT bEnable) OR _bFault THEN
        _eState := E_DL_N2PurgeState.eFault;         // 失能或故障：进故障相
    ELSIF NOT _bInBand THEN
        IF tonEstablish.Q THEN
            _bEstTimeout := TRUE;                    // 吹扫中流量持续离带：按建立失败处理
            _uFault := 16#0003_021F;                 // 故障级：建立超时（复用同一根因码）
            _bFault := TRUE;                         // 锁存
            bError  := TRUE;                         // 故障标志置位（R45 配对）
            _eState := E_DL_N2PurgeState.eTimeout;   // 进超时相
        END_IF
    ELSIF rtStart.Q THEN
        _bEstBreak := TRUE;                          // 再次起始：重建窗口（不停吹扫）
        _bInBandBrk := TRUE;                         // 入带计时重启
    END_IF

E_DL_N2PurgeState.eTimeout:
    IF (NOT _bFault) AND (NOT _bCfgBad) AND bEnable AND _bInBand THEN
        _eState := E_DL_N2PurgeState.ePurged;        // 流量恢复入带且码已清：回吹扫相
        _bEstTimeout := FALSE;                       // 超时保持量释放（与按码专清同源）
    END_IF

E_DL_N2PurgeState.eFault:
    IF (NOT _bFault) AND (NOT _bCfgBad) AND bEnable THEN
        _eState := E_DL_N2PurgeState.eIdle;          // 锁存已清且组态合法：回空闲等下一次起始
    END_IF

ELSE
    _uFault := 16#0003_025F;                         // 故障级：相位 ID 越界（枚举兜底）
    _bFault := TRUE;                                 // 锁存
    bError  := TRUE;                                 // 故障标志置位（R45 配对）
    _eState := E_DL_N2PurgeState.eFault;             // 强制回故障相
END_CASE

(* 段 5B｜021F 按码专清：入带持续窗满且无其它故障 → 建立超时可解（R188 可达清除边） *)
IF (_uFault = 16#0003_021F) AND _bInBand AND tonInBand.Q THEN
    _uFault := 16#0000_0000;                         // 清锁存码
    _bFault := FALSE;                                // 锁存位同步清
    _bEstTimeout := FALSE;                           // 超时保持量与码同源释放
END_IF

(* —— 段 6：故障码优先级链（信号无效优先于越限，越限优先于超时；R190 归因唯一） —— *)
IF _bCfgBad THEN
    _uFault := 16#0003_020F;                         // 组态非法优先上报
    _bFault := TRUE;
    bError  := TRUE;
ELSIF _bDewBad THEN
    _uFault := 16#0003_022F;                         // 露点信号无效优先于数值判据
    _bFault := TRUE;
    bError  := TRUE;
END_IF

(* —— 段 7：出口单点映射（名实同源；锁存码回放，禁同拍抹除） —— *)
bEstablishTimeout := _bEstTimeout;                   // 建立超时出口（保持型）
bDewPointAlarm    := _bDewAlarm;                     // 露点越限出口（保持型）
bDewSevereAlarm   := _bDewSevere;                    // 严重越限出口（保持型）
bPurgeOk := bEnable AND (_eState = E_DL_N2PurgeState.ePurged) AND _bInBand AND
            (NOT _bDewAlarm) AND (NOT _bDewBad) AND (NOT _bFault) AND (NOT _bCfgBad);  // 合格判定（全条件）
eStateOut := _eState;                                // 状态出口
IF _bFault THEN
    nErrId := _uFault;                               // 故障锁存码回放（不在故障相按当下输入重推）
    bError := TRUE;                                  // 故障出口派生自锁存
ELSE
    nErrId := _uInfo;                                // 信息码
END_IF
bValid := bEnable AND (NOT _bFault) AND (NOT _bCfgBad);  // 判据可用

END_FUNCTION_BLOCK

(* ---- FB_DL_FreshAirStepperDamper.st ---- *)
(*
  FB_DL_FreshAirStepperDamper  —  新风阀步进执行器开环驱动 / Fresh-air stepper damper open-loop driver
  分类 Category : DL_Device
  码位 Code     : 16#03_2_16
  段位说明      : 03_2 段低半字节 00~0F 已满（05 为历史空穴留存），进位 16 段续号（R192）
  版本 Version  : 1.0.0
  来源 Source   : t1-2-oscat-building — IEC 61131-3 标准语义的道莅防御性实现
  溯源 Origin   : OSCAT 楼控步进阀公开语义借鉴，clean-room 实现，未复制任何源码行
                  （与 FB_DL_PulseDirStepper 分工：本件带开度当量换算与端点自学习；裸脉冲/方向驱动由 PulseDirStepper 承载）
  功能 Function : 1) 开度↔步数当量换算：目标步数 = fOpenCmdPct/100 × nStepsFullStroke，经 iStepper.MoveRelative 单发下发；
                  2) 反向行进时额外补 nBacklashSteps 间隙步（同向不补，间隙单向补偿）；
                  3) 端点自学习：回零撞负限位（uAlarmWord bit1）或超步数判 bAtEndStop 后清计数定标；
                  4) 未回零拒绝开度指令（只允许回零，置信息码）。
  边界 Boundary : ① nStepsFullStroke <= 0 / fStepRateHz <= 0 防除零判组态错；
                  ② fOpenCmdPct 越 0~100 钳制并置信息码；nBacklashSteps < 0 取 ABS 并置信息码；
                  ③ 位置计数 DINT 且到 [0, nStepsFullStroke] 边界钳制禁回绕（R28-2 两点向量：0% 计数钳 0 不出负值；
                     100% 计数钳 nStepsFullStroke 不越上界）；
                  ④ 步进接口按「步当量」下发（1 当量 = 1 步），单位换算由上层适配层承载；
                  ⑤ 解除式自证：bAtEndStop 解除 = 离开端点的 MoveRelative 受理（定标后计数已清零）；
                  ⑥ CASE 全态覆盖 + ELSE 兜底置故障相。
  依赖 Depends  : I_DL_StepperOpenLoop（注入，不实例化）；语义对齐 FB_DL_ToleranceWindow（已注册，不实例化）
  码表 Error codes（本件格 03_2_16，子码步进 +0x100）:
    16#0003_0116 信息级：未回零拒开度指令（只允许回零）
    16#0003_0216 故障级：组态非法（全行程步数 <= 0 / 步频 <= 0），锁存至复位
    16#0003_0316 信息级：开度越 0..100 已钳制
    16#0003_0416 信息级：反向间隙步数为负，已取 ABS
    16#0003_0516 信息级：端点定标完成（计数清零）
    16#0003_0616 故障级：状态机落 ELSE 兜底（非法相位 ID）

  修订历史 Revision :
    2026-11-18  v1.0.0  R38 首版
*)

TYPE E_DL_DamperState :
(
    eUnhomed := 0,    // 未回零：只允许回零指令 / Unhomed, only homing allowed
    eHoming  := 10,   // 回零中：向端点步进 / Homing, stepping toward end stop
    eReady   := 20,   // 就绪：已定标待机 / Ready, calibrated and idle
    eMoving  := 30,   // 行进中：开度指令执行中 / Moving, executing position command
    eFault   := 90    // 故障：组态/驱动故障锁定 / Fault, latched
);
END_TYPE

FUNCTION_BLOCK FB_DL_FreshAirStepperDamper
VAR_INPUT
    fOpenCmdPct     : REAL := 0.0;       // 开度指令 [%]，域 0..100 / Open command percentage
    bHomingCmd      : BOOL := FALSE;     // 回零指令 / Homing command
    nStepsFullStroke: INT  := 1000;      // 全行程步数 [步]，域 > 0 / Full-stroke step count
    nBacklashSteps  : INT  := 5;         // 反向间隙步数 [步]，< 0 取 ABS / Backlash steps
    fStepRateHz     : REAL := 200.0;     // 步进频率 [Hz]，域 > 0 / Step rate
    bReset          : BOOL := FALSE;     // 复位（Fault 解除路径）/ Reset
END_VAR
VAR_OUTPUT
    fActualPosPct   : REAL;              // 实际开度 [%]（开环推算）/ Actual open percentage
    nStepCount      : DINT;              // 位置步计数 [步]，域 [0, 全行程] / Position step count
    bHoming         : BOOL;              // 回零进行中 / Homing in progress
    bHomed          : BOOL;              // 已回零定标 / Homed flag
    bAtEndStop      : BOOL;              // 端点判据成立 / At end stop
    nErrId          : UDINT;             // 事件码，0 = 无事件 / Event code
    eState          : E_DL_DamperState;  // 状态出口，段尾单点映射 / State outlet
END_VAR
VAR_IN_OUT
    iStepper : I_DL_StepperOpenLoop;     // 步进执行器引用（注入，不实例化）/ Stepper reference, injected
END_VAR
VAR
    tonReadyWch : TON;                   // 受理回读观察窗（单发后等 bReady），自复位 / Acceptance watch window
    tonFaultWch : TON;                   // 故障观察窗，自复位 / Fault watch window, self-resetting
    rtHome      : R_TRIG;                // 回零指令上升沿 / Homing command rising edge
    rtReset     : R_TRIG;                // 复位上升沿 / Reset rising edge
    _eState     : E_DL_DamperState := E_DL_DamperState.eUnhomed;   // 内部相位（CASE 唯一写入目标）/ Internal phase
    _nTarget    : INT;                   // 目标步数 [步] / Target step count
    _nDelta     : INT;                   // 本拍步增量 [步] / Step delta this scan
    _nBlCmp     : INT;                   // 间隙补偿生效步数 [步] / Effective backlash compensation
    _rClampCmd  : REAL;                  // 钳制后开度指令 [%] / Clamped open command
    _uFault     : UDINT;                 // 故障码锁存 / Latched fault code
    _uInfo      : UDINT;                 // 信息码，每拍重算 / Info code
    _bFault     : BOOL;                  // 故障锁存位 / Latched fault bit
    _bCfgBad    : BOOL;                  // 组态非法聚合 / Configuration invalid aggregate
    _bCmdPend   : BOOL;                  // 单发待受理标志 / One-shot pending acceptance flag
    _bHomePend  : BOOL;                  // 回零单发待受理标志 / Homing one-shot pending flag
    _nHomeSteps : INT;                   // 回零行程步数（含裕度）[步] / Homing travel steps with margin
END_VAR
VAR CONSTANT
    DL_ALM_NEG_LIM : WORD := 16#0002;    // 报警字 bit1 负限位 / Alarm word bit1 negative limit
    DL_HOME_MARGIN : INT  := 50;         // 回零裕度步数 [步] / Homing margin steps
    DL_WATCH_PT    : TIME := T#2S;       // 故障观察窗 [ms]，自复位 / Fault watch window
    DL_READY_PT    : TIME := T#5S;       // 受理回读观察窗 [ms] / Acceptance watch window
END_VAR

(* —— 段 0：定时器与边沿无条件周期刷新（R182：调用语句不得置于 IF/CASE 内） —— *)
rtHome(CLK := bHomingCmd);                                       // 回零上升沿，每拍必调
rtReset(CLK := bReset);                                          // 复位上升沿，每拍必调
tonFaultWch(IN := (NOT tonFaultWch.Q), PT := DL_WATCH_PT);       // 观察窗自复位（表达式入参）
tonReadyWch(IN := _bCmdPend OR _bHomePend, PT := DL_READY_PT);   // 受理回读观察窗（表达式入参）

(* —— 段 1：单拍量预清零（锁存量 _uFault/_bFault/_nStepCount/_bHomed 不入清单，R187①） —— *)
_uInfo := 16#0000_0000;         // 信息码每拍重算
bHoming := FALSE;               // 回零出口缺省 FALSE（段 8 单点置位）
bAtEndStop := FALSE;            // 端点出口缺省 FALSE（Homing 相单点置位）
_bCfgBad := FALSE;              // 组态非法预清零
nErrId := 16#0000_0000;         // 事件码缺省无事件

(* —— 段 2：组态域闸（覆盖全部参与判据换算的引脚，R151） —— *)
IF (nStepsFullStroke <= 0) OR (fStepRateHz <> fStepRateHz) OR (fStepRateHz <= 0.0) THEN
    _bCfgBad := TRUE;           // 全行程步数/步频非法（防除零）
END_IF

(* —— 段 3：复位沿（Fault 解除唯一路径：bReset） —— *)
IF rtReset.Q THEN
    _bFault := FALSE;           // 清故障锁存位
    _uFault := 16#0000_0000;
    _bCmdPend := FALSE;         // 受理标志复位
    _bHomePend := FALSE;
    _eState := E_DL_DamperState.eUnhomed;   // 复位回未回零（定标状态重判）
END_IF

(* —— 段 4：输入归一（钳制 + 间隙 ABS，均置信息码） —— *)
IF fOpenCmdPct < 0.0 THEN
    _rClampCmd := 0.0;          // 越下限钳 0（R28-2 向量一：0% 不回绕负值）
    _uInfo := 16#0003_0316;     // 信息级：开度越域已钳制
ELSIF fOpenCmdPct > 100.0 THEN
    _rClampCmd := 100.0;        // 越上限钳 100（R28-2 向量二：100% 不越上界）
    _uInfo := 16#0003_0316;     // 信息级：开度越域已钳制
ELSE
    _rClampCmd := fOpenCmdPct;  // 域内直通
END_IF
IF nBacklashSteps < 0 THEN
    _nBlCmp := -nBacklashSteps; // 负间隙步取 ABS（规格强制）
    _uInfo := 16#0003_0416;     // 信息级：负间隙步已取 ABS
ELSE
    _nBlCmp := nBacklashSteps;  // 正常值直通
END_IF
_nTarget := TRUNC(_rClampCmd / 100.0 * INT_TO_REAL(nStepsFullStroke));   // 开度→步数当量换算

(* —— 段 5：相位机（只做迁移与单发命令；出口在段 8） —— *)
CASE _eState OF

E_DL_DamperState.eUnhomed:
    IF _bCfgBad THEN
        _uFault := 16#0003_0216;            // 故障级：组态非法
        _bFault := TRUE;                    // 锁存（复位沿可清）
        _eState := E_DL_DamperState.eFault;
    ELSIF rtHome.Q THEN
        _nHomeSteps := nStepsFullStroke + _nBlCmp + DL_HOME_MARGIN;   // 回零行程（含裕度）
        iStepper.MoveRelative(fDistance := INT_TO_LREAL(-_nHomeSteps), fSpeed := fStepRateHz);   // 单发向端点
        _bHomePend := TRUE;                 // 待受理标志
        _eState := E_DL_DamperState.eHoming;// 进回零相
    ELSIF _nTarget <> DINT_TO_INT(nStepCount) THEN
        _uInfo := 16#0003_0116;             // 信息级：未回零拒开度指令（只允许回零）
    END_IF

E_DL_DamperState.eHoming:
    bAtEndStop := (iStepper.uAlarmWord AND DL_ALM_NEG_LIM) <> 0;   // 端点判据：负限位报警字
    IF bAtEndStop OR tonReadyWch.Q THEN
        nStepCount := 0;                    // 端点定标：计数清零（禁回绕）
        bHomed := TRUE;                     // 定标完成
        _uInfo := 16#0003_0516;             // 信息级：端点定标完成
        _bHomePend := FALSE;                // 受理标志清
        _eState := E_DL_DamperState.eReady; // 进就绪相
    ELSIF iStepper.uAlarmWord <> 0 THEN
        IF (iStepper.uAlarmWord AND DL_ALM_NEG_LIM) = 0 THEN
            _uFault := 16#0003_0216;        // 回零中出现非限位报警（驱动器/堵转）：按组态域故障升级
            _bFault := TRUE;
            iStepper.Stop();
            _eState := E_DL_DamperState.eFault;
        END_IF
    END_IF

E_DL_DamperState.eReady:
    IF _nTarget <> DINT_TO_INT(nStepCount) THEN
        _nDelta := _nTarget - DINT_TO_INT(nStepCount);              // 步增量
        IF (_nDelta < 0) AND (_nBlCmp > 0) THEN
            _nDelta := _nDelta - _nBlCmp;                           // 反向行进：额外补间隙步（同向不补）
        END_IF
        iStepper.MoveRelative(fDistance := INT_TO_LREAL(_nDelta), fSpeed := fStepRateHz);   // 单发下发（步当量）
        nStepCount := DINT(_nTarget);                               // 开环指令位置记账（钳制见段 6）
        _bCmdPend := TRUE;                                          // 待受理标志
        _eState := E_DL_DamperState.eMoving;                        // 进行进相
    ELSIF iStepper.uAlarmWord <> 0 THEN
        _uFault := 16#0003_0216;            // 就绪态出现驱动报警
        _bFault := TRUE;
        _eState := E_DL_DamperState.eFault;
    END_IF

E_DL_DamperState.eMoving:
    IF iStepper.bReady THEN
        _bCmdPend := FALSE;                 // 受理确认
        _eState := E_DL_DamperState.eReady; // 回就绪相
    ELSIF tonReadyWch.Q THEN
        _uFault := 16#0003_0216;            // 受理回读超观察窗（驱动无响应）
        _bFault := TRUE;
        iStepper.Stop();
        _eState := E_DL_DamperState.eFault;
    ELSIF iStepper.uAlarmWord <> 0 THEN
        _uFault := 16#0003_0216;            // 行进中出现驱动报警
        _bFault := TRUE;
        iStepper.Stop();
        _eState := E_DL_DamperState.eFault;
    END_IF

E_DL_DamperState.eFault:
    ;                                       // 故障相：等复位沿（段 3 承载解除）

ELSE
    _uFault := 16#0003_0616;                // 故障级：非法相位 ID 兜底
    _bFault := TRUE;                        // 锁存
    _eState := E_DL_DamperState.eFault;     // 强制回故障相

END_CASE

(* —— 段 6：位置计数边界钳制（禁回绕，R28-2 两点向量收口） —— *)
IF nStepCount < 0 THEN
    nStepCount := 0;                        // 下界钳 0（0% 向量：不出负计数）
ELSIF nStepCount > DINT(nStepsFullStroke) THEN
    nStepCount := DINT(nStepsFullStroke);   // 上界钳全行程（100% 向量：不越上界）
END_IF

(* —— 段 7：出口单点映射（名实同源；锁存码回放，禁同拍抹除） —— *)
fActualPosPct := DINT_TO_REAL(nStepCount) * 100.0 / INT_TO_REAL(nStepsFullStroke);   // 开度出口（分母已闸 > 0）
bHoming := (_eState = E_DL_DamperState.eHoming);          // 回零出口（相位单点）
bHomed := bHomed AND (NOT _bFault);       // 定标出口（故障相撤销）
bAtEndStop := bAtEndStop AND (_eState = E_DL_DamperState.eHoming);   // 端点出口仅回零相有效
IF _bFault THEN
    nErrId := _uFault;          // 故障锁存码回放
ELSIF _uInfo <> 16#0000_0000 THEN
    nErrId := _uInfo;           // 信息码
END_IF
eState := _eState;              // 状态出口单点映射

END_FUNCTION_BLOCK

(* ---- FB_DL_FrostProtectFreeze.st ---- *)
(*==============================================================================
 * 组件名称 (Component)  : FB_DL_FrostProtectFreeze
 * 所属子库 (Sublibrary) : DL_Device
 * 当前版本 (Version)    : 1.0.0
 * 兼容性 (Platform)     : CODESYS 3.5 / TwinCAT 3 / 汇川 InoProShop / Machine Expert
 *                         仅依赖纯 IEC 61131-3 标准元素，零厂商方言
 * 功能描述 (Function)   : 防冻保护：委托 FC_DL_Hysteresis 双阈判定（设定 ± 回差）
 *                         联动新风阀关闭 / 盘管阀开 + 风机停机；NORMAL → WARN →
 *                         TRIP（三输出同拍安全态）→ 人工复位 → RESET（条件核实）→
 *                         NORMAL。TRIP 后必须 bManualReset 才退出（安全侧保持）。
 * 溯源 (Origin)         : 道莅 clean-room 防御性实现
 * 本文件内含 (Contains) : TYPE E_DL_FrostState / TYPE E_DL_FrostErr /
 *                         FUNCTION_BLOCK FB_DL_FrostProtectFreeze
 * 依赖 (Depends)        : DL_MathData/FC_DL_Hysteresis
 * 红线自检 (Redline)    : 无外部全局变量、无硬件地址直引 ｜ 全变量中英双语同行注释
 *                         非有限值防御 + 量程钳位 + 回差下限钳制 ｜ 枚举成员全部显式赋值
 *                         状态机 CASE 含 ELSE 兜底（ELSE → 安全态输出）｜ 无定时器实例
 * 错误码表 (Codes)      : 16#0003_0393 NORMAL
 *                         16#0003_0394 WARN（接近防冻设定）
 *                         16#0003_0395 TRIP(冻结输出保持)
 *                         16#0003_0396 复位挂起(恢复条件未满足)
 *                         16#0003_0397 传感器无效(保持上次安全态)
 * 修订历史 (Revision)   : 2026-11-17  v1.0.0  首版入库 · R27 · 阶段三批 2
 * 验收向量 (Acceptance) : 设定 4 C 回差 1 C：室外 3.0 → TRIP；室外 5.5+复位 → RESET→NORMAL；
 *                         bFrostAlarm=TRUE → 直进 TRIP；温度 NaN → 0397 保持安全态
 *============================================================================*)

(*-----------------------------------------------------------------------------
 * 枚举: E_DL_FrostState（归属 DL_Device，防冻状态机状态）
 *----------------------------------------------------------------------------*)
TYPE E_DL_FrostState :
(
    eNormal := 0,    // 正常：防冻判据未触发 / Normal, no frost trip
    eWarn   := 10,   // 预警：温度接近防冻设定（迟滞带内）/ Warning, temperature near the setpoint
    eTrip   := 20,   // 跳闸：防冻触发，三输出安全态保持 / Tripped, safe outputs held
    eReset  := 30,   // 复位挂起：人工已复位但恢复条件未核实 / Reset pending, conditions unverified
    eFault  := 99    // 传感器无效兜底态 / Sensor-invalid fallback
);
END_TYPE

(*-----------------------------------------------------------------------------
 * 枚举: E_DL_FrostErr（归属 DL_Device，与 FB_DL_FrostProtectFreeze 同文件）
 *----------------------------------------------------------------------------*)
TYPE E_DL_FrostErr :
(
    eNormal    := 16#0003_0393,   // NORMAL / Normal
    eWarn      := 16#0003_0394,   // WARN（接近防冻设定）/ Warning near setpoint
    eTrip      := 16#0003_0395,   // TRIP（冻结输出保持）/ Tripped, outputs held
    eResetHold := 16#0003_0396,   // 复位挂起（条件未满足）/ Reset pending
    eSensorBad := 16#0003_0397    // 传感器无效（保持上次安全态）/ Sensor invalid
);
END_TYPE

(*==============================================================================
 * 功能块: FB_DL_FrostProtectFreeze
 * 调用约定: 每个扫描周期无条件调用一次。
 *============================================================================*)
FUNCTION_BLOCK FB_DL_FrostProtectFreeze
VAR_INPUT
    fFrostTemp_C  : REAL;              // 防冻温度设定 [摄氏度]，默认 4 / Frost protection setpoint [degC]
    fOutdoor_C    : REAL;              // 室外温度 [摄氏度]，有效域 -50~60 / Outdoor temperature [degC]
    bHysteresisC  : REAL;              // 回差 [摄氏度]，默认 1.0，下限钳 0.1 / Hysteresis width [degC]
    bFrostAlarm   : BOOL;              // 盘管防冻开关输入（硬件低温断路器）/ Coil frost switch input
    bManualReset  : BOOL;              // 人工复位（TRIP 退出门票）/ Manual reset, trip exit ticket
END_VAR
VAR_OUTPUT
    bDamperCloseCmd : BOOL;            // 关新风阀指令 / Damper close command
    bCoilOpenCmd    : BOOL;            // 开盘管阀指令 / Coil valve open command
    bFanStopCmd     : BOOL;            // 风机停机指令 / Fan stop command
    eState          : E_DL_FrostState; // 防冻状态机当前状态 / Frost state machine state
    eErr            : E_DL_FrostErr;   // 错误码 / Error code
END_VAR
VAR
    bHystState   : BOOL;               // 迟滞状态（调用方持有并回传）/ Hysteresis state held by caller
    fTempUse     : REAL;               // 生效室外温度（钳位后）[摄氏度] / Effective outdoor temperature [degC]
    fSetUse      : REAL;               // 生效设定（NaN 兜底）[摄氏度] / Effective setpoint [degC]
    fHystUse     : REAL;               // 生效回差（钳位后）[摄氏度] / Effective hysteresis [degC]
    bFrostTrip   : BOOL;               // 防冻跳闸判据（迟滞+开关合成）/ Frost trip predicate
    bNonFin      : BOOL;               // 非有限输入汇总标志 / Non-finite input aggregate flag
    uHystErr     : UDINT;              // 委托迟滞错误码（0 = 无错）/ Delegate hysteresis error id
    fUpTrip      : REAL;               // 委托输出：实际上阈值 [摄氏度] / Delegate upper trip [degC]
    fLoTrip      : REAL;               // 委托输出：实际下阈值 [摄氏度] / Delegate lower trip [degC]
END_VAR
VAR CONSTANT
    DL_FRS_T_MIN    : REAL := -50.0;   // 室外温度域下限 [摄氏度] / Outdoor temperature lower bound [degC]
    DL_FRS_T_MAX    : REAL := 60.0;    // 室外温度域上限 [摄氏度] / Outdoor temperature upper bound [degC]
    DL_FRS_HYST_MIN : REAL := 0.1;     // 回差下限 [摄氏度] / Hysteresis lower bound [degC]
    DL_FRS_SET_DFLT : REAL := 4.0;     // 设定兜底值 [摄氏度] / Setpoint fallback [degC]
    DL_FRS_INF_MAX  : REAL := 1.0E30;  // 非有限值判定幅值上限 / Magnitude bound for finite-value check
    DL_FRS_ZERO     : REAL := 0.0;     // 零值常量，避免裸字面量 / Zero constant
END_VAR

(*------------------------------------------------------------------------------
 * 段 1｜非有限值闸：设定/温度 NaN 或溢出 → 0397 保持安全态输出
 *----------------------------------------------------------------------------*)
bNonFin := (fFrostTemp_C <> fFrostTemp_C) OR (ABS(fFrostTemp_C) > DL_FRS_INF_MAX)
        OR (fOutdoor_C    <> fOutdoor_C)    OR (ABS(fOutdoor_C)    > DL_FRS_INF_MAX)
        OR (bHysteresisC  <> bHysteresisC)  OR (ABS(bHysteresisC)  > DL_FRS_INF_MAX);
IF bNonFin THEN
    eState := E_DL_FrostState.eFault;                // 进传感器无效兜底态 / enter sensor-invalid fallback
    eErr := E_DL_FrostErr.eSensorBad;                // 信息级：传感器无效 / sensor invalid
    bDamperCloseCmd := TRUE;                         // 安全态：关新风阀 / safe: close damper
    bCoilOpenCmd := TRUE;                            // 安全态：开盘管阀 / safe: open coil valve
    bFanStopCmd := TRUE;                             // 安全态：风机停机 / safe: stop fan
    RETURN;
END_IF

(*------------------------------------------------------------------------------
 * 段 2｜参数钳位：室外温 [-50,60]、回差下限 0.1、设定兜底
 *----------------------------------------------------------------------------*)
fTempUse := fOutdoor_C;                              // 温度工作副本 / temperature working copy
IF fTempUse < DL_FRS_T_MIN THEN
    fTempUse := DL_FRS_T_MIN;                        // 下限钳位 / floored
ELSIF fTempUse > DL_FRS_T_MAX THEN
    fTempUse := DL_FRS_T_MAX;                        // 上限钳位 / capped
END_IF
fSetUse := fFrostTemp_C;                             // 设定工作副本 / setpoint working copy
IF (fSetUse <= DL_FRS_T_MIN) OR (fSetUse >= DL_FRS_T_MAX) THEN
    fSetUse := DL_FRS_SET_DFLT;                      // 设定出域按兜底值（配置防御）/ setpoint out of domain falls back
END_IF
fHystUse := bHysteresisC;                            // 回差工作副本 / hysteresis working copy
IF fHystUse < DL_FRS_HYST_MIN THEN
    fHystUse := DL_FRS_HYST_MIN;                     // 回差下限钳位 / hysteresis floored
END_IF

(*------------------------------------------------------------------------------
 * 段 3｜委托迟滞双阈判定（FC_DL_Hysteresis，状态由本块持有回传）
 *----------------------------------------------------------------------------*)
FC_DL_Hysteresis(fIn := fTempUse, fThreshold := fSetUse, fHysteresis := fHystUse,
                 bState := bHystState, fUpperTrip => fUpTrip, fLowerTrip => fLoTrip,
                 uErrorId => uHystErr);              // 迟滞委托：bHystState 为 TRUE 表示温度低于下阈 / delegate: TRUE means below lower trip
bFrostTrip := bHystState OR bFrostAlarm;             // 跳闸判据 = 迟滞触发或硬件开关 / trip predicate

(*------------------------------------------------------------------------------
 * 段 4｜状态机：CASE 含 ELSE 兜底（ELSE → 安全态输出）
 *----------------------------------------------------------------------------*)
CASE eState OF

    E_DL_FrostState.eNormal:
        bDamperCloseCmd := FALSE;                    // 正常态不关阀 / no damper close in normal
        bCoilOpenCmd := FALSE;                       // 正常态不开盘管阀 / no coil valve in normal
        bFanStopCmd := FALSE;                        // 正常态不停风机 / no fan stop in normal
        IF fTempUse < (fSetUse - fHystUse) THEN
            eState := E_DL_FrostState.eWarn;         // 接近设定：预警 / near setpoint: warning
        END_IF
        IF bFrostTrip THEN
            eState := E_DL_FrostState.eTrip;         // 跳闸判据成立：直进 TRIP / trip predicate: enter trip
        END_IF

    E_DL_FrostState.eWarn:
        bDamperCloseCmd := FALSE;                    // 预警不动作（仅提示）/ warning only, no action
        bCoilOpenCmd := FALSE;                       // 预警不动作 / no action on warning
        bFanStopCmd := FALSE;                        // 预警不动作 / no action on warning
        IF bFrostTrip THEN
            eState := E_DL_FrostState.eTrip;         // 跳闸判据成立：TRIP / trip predicate: enter trip
        ELSIF fTempUse > fSetUse THEN
            eState := E_DL_FrostState.eNormal;       // 温度回升过设定：回正常 / recovered above setpoint
        END_IF

    E_DL_FrostState.eTrip:
        bDamperCloseCmd := TRUE;                     // TRIP 安全态：关新风阀 / trip safe: close damper
        bCoilOpenCmd := TRUE;                        // TRIP 安全态：开盘管阀 / trip safe: open coil valve
        bFanStopCmd := TRUE;                         // TRIP 安全态：风机停机 / trip safe: stop fan
        IF bManualReset THEN
            eState := E_DL_FrostState.eReset;        // 人工复位进核实相 / manual reset enters reset-pending
        END_IF

    E_DL_FrostState.eReset:
        bDamperCloseCmd := TRUE;                     // 核实相保持安全态（条件未满足不撤）/ safe outputs held while unverified
        bCoilOpenCmd := TRUE;                        // 核实相保持安全态 / safe outputs held
        bFanStopCmd := TRUE;                         // 核实相保持安全态 / safe outputs held
        IF bFrostTrip THEN
            eState := E_DL_FrostState.eTrip;         // 跳闸判据仍在：退回 TRIP / predicate persists: back to trip
        ELSIF (NOT bFrostTrip) AND (fTempUse > fSetUse) THEN
            eState := E_DL_FrostState.eNormal;       // 恢复条件满足（温度过设定且开关释放）/ recovery conditions met
        ELSE
            eState := E_DL_FrostState.eReset;        // 条件未满足：复位挂起 / conditions unmet, reset pending
        END_IF

    E_DL_FrostState.eFault:
        bDamperCloseCmd := TRUE;                     // 兜底态保持安全输出 / fallback holds safe outputs
        bCoilOpenCmd := TRUE;                        // 兜底态保持安全输出 / fallback holds safe outputs
        bFanStopCmd := TRUE;                         // 兜底态保持安全输出 / fallback holds safe outputs
        IF (NOT bNonFin) THEN
            eState := E_DL_FrostState.eNormal;       // 输入恢复有限后自动回正常（传感器无效不锁存）/ auto-recover when input finite again
        END_IF

    ELSE
        eState := E_DL_FrostState.eFault;            // 非法状态兜底 / illegal-state fallback
        eErr := E_DL_FrostErr.eSensorBad;            // 兜底码（传感器无效段，反证句：输出同为三安全态）/ fallback code
        bDamperCloseCmd := TRUE;                     // 安全态输出 / safe outputs
        bCoilOpenCmd := TRUE;                        // 安全态输出 / safe outputs
        bFanStopCmd := TRUE;                         // 安全态输出 / safe outputs

END_CASE

(*------------------------------------------------------------------------------
 * 段 5｜状态码映射（信息级状态码随状态输出）
 *----------------------------------------------------------------------------*)
CASE eState OF
    E_DL_FrostState.eNormal:
        eErr := E_DL_FrostErr.eNormal;               // 码 0393 / code normal
    E_DL_FrostState.eWarn:
        eErr := E_DL_FrostErr.eWarn;                 // 码 0394 / code warn
    E_DL_FrostState.eTrip:
        eErr := E_DL_FrostErr.eTrip;                 // 码 0395 / code trip
    E_DL_FrostState.eReset:
        eErr := E_DL_FrostErr.eResetHold;            // 码 0396 / code reset pending
    E_DL_FrostState.eFault:
        eErr := E_DL_FrostErr.eSensorBad;            // 码 0397 / code sensor invalid
    ELSE
        eErr := E_DL_FrostErr.eSensorBad;            // 非法状态兜底码 / illegal-state fallback code
END_CASE
END_FUNCTION_BLOCK

(* ---- FB_DL_FurnaceBeltTension.st ---- *)
// =====================================================================
// FB_DL_FurnaceBeltTension.st
// 烧结炉网带张力闭环 + 边缘跑偏纠偏（双环加权共用执行器）
// Furnace belt tension loop + edge steering FB
// 码位: 16#0003_03D4 ~ 16#0003_03D8 (本件独占 5 槽)
// 修改记录: R29 初版 (按 DISPATCH_R29 序 11)
// =====================================================================
FUNCTION_BLOCK FB_DL_FurnaceBeltTension
VAR_INPUT
    bEnable        : BOOL  := FALSE;   // 使能 / Enable
    bWebRun        : BOOL  := FALSE;   // 网带运行 / Web running
    fTension_N     : REAL  := 0.0;     // 实测张力 0~5000 N / Measured tension [N]
    fTensionSp_N   : REAL  := 800.0;   // 张力设定 0~5000 N / Tension setpoint [N]
    fEdgePos_mm    : REAL  := 0.0;     // 边缘位置 -50~50 mm（正=右偏）/ Edge position [mm]
    fEdgeCenter_mm : REAL  := 0.0;     // 边缘中心基准 -50~50 mm / Edge center [mm]
    fEdgeTol_mm    : REAL  := 3.0;     // 跑偏容差 0.1~20 mm / Edge tolerance [mm]
    fTensionTolPct : REAL  := 5.0;     // 张力容差 0.5~50 % / Tension tolerance [%]
    fKpT           : REAL  := 0.02;    // 张力环增益 0.001~1 %/N / Tension gain [%/N]
    fKpE           : REAL  := 0.5;     // 纠偏环增益 0.01~5 %/mm / Edge gain [%/mm]
    fTrimMax_pct   : REAL  := 10.0;    // 输出限幅 0.5~50 % / Output limit [%]
    fWeightT       : REAL  := 0.7;     // 张力权重 0~1 / Tension weight [-]
END_VAR
VAR_OUTPUT
    fTrimOut_pct   : REAL;              // 速度微调 -100~100 % / Speed trim [%]
    fDev_N         : REAL;              // 张力偏差 N / Tension deviation [N]
    fEdgeDev_mm    : REAL;              // 边缘偏差 mm / Edge deviation [mm]
    bTensionAlarm  : BOOL;              // 张力超差 / Tension alarm
    bEdgeAlarm     : BOOL;              // 跑偏超差 / Edge alarm
    eErr           : UDINT;             // 错误码 / Error code
END_VAR
VAR
    fWeightTSafe   : REAL;              // 钳 [0,1] 后张力权重 / Clamped tension weight [-]
    fWeightE       : REAL;              // 纠偏权重 = 1-张力权重 / Edge weight [-]
    fTensionTrim   : REAL;              // 张力环输出项 / Tension loop term [%]
    fEdgeTrim      : REAL;              // 纠偏环输出项 / Edge loop term [%]
    fTolPctSafe    : REAL;              // 张力容差处理值 / Sanitized tension tolerance [%]
    fEdgeTolSafe   : REAL;              // 跑偏容差处理值 / Sanitized edge tolerance [mm]
    bSatLatch      : BOOL := FALSE;     // 饱和故障锁存 / Saturation fault latch
    tonSat         : TON;               // 饱和持续计时（无条件刷新）/ Saturation timer
    bSatCond       : BOOL;              // 饱和条件当前值 / Saturation condition
    xFirstScan     : BOOL  := TRUE;     // 首扫标记 / First-scan flag
END_VAR

// ---------------------------------------------------------------------
// 代码位表（本件独占，勿复用）:
//   16#0003_03D4 信息 双环运行正常
//   16#0003_03D5 故障 输入非有限
//   16#0003_03D6 故障 fTensionSp_N ≤ 0 / fTrimMax_pct ≤ 0 / fKpT ≤ 0 / fKpE < 0（组态错）；fEdgeTol ≤ 0 兜底登记同槽
//   16#0003_03D7 信息 bWebRun=FALSE 或 bEdgeAlarm=TRUE → 输出归 0 / 张力环冻结，积分保持
//   16#0003_03D8 故障 张力环输出持续 10 s 触限仍同向偏差 > 容差 → 锁存，解除需 bReset
// ---------------------------------------------------------------------

// ---- 非有限闸 / Finite gate ----
IF (fTension_N <> fTension_N) OR (ABS(fTension_N) >= 1.0E12)
   OR (fTensionSp_N <> fTensionSp_N) OR (ABS(fTensionSp_N) >= 1.0E12)
   OR (fEdgePos_mm <> fEdgePos_mm) OR (ABS(fEdgePos_mm) >= 1.0E12)
   OR (fEdgeCenter_mm <> fEdgeCenter_mm) OR (ABS(fEdgeCenter_mm) >= 1.0E12)
   OR (fEdgeTol_mm <> fEdgeTol_mm) OR (ABS(fEdgeTol_mm) >= 1.0E12)
   OR (fTensionTolPct <> fTensionTolPct) OR (ABS(fTensionTolPct) >= 1.0E12)
   OR (fKpT <> fKpT) OR (ABS(fKpT) >= 1.0E12)
   OR (fKpE <> fKpE) OR (ABS(fKpE) >= 1.0E12)
   OR (fTrimMax_pct <> fTrimMax_pct) OR (ABS(fTrimMax_pct) >= 1.0E12)
   OR (fWeightT <> fWeightT) OR (ABS(fWeightT) >= 1.0E12) THEN
    fTrimOut_pct := 0.0;        // 输出归 0（安全侧）/ Output zero
    bTensionAlarm := FALSE;     // 报警复位 / Alarm reset
    eErr := 16#0003_03D5;       // 故障码 / Fault code
    RETURN;                     // 本拍结束 / End of cycle
END_IF

// ---- 组态错闸 / Configuration fault gate ----
IF (fTensionSp_N <= 0.0) OR (fTrimMax_pct <= 0.0) OR (fKpT <= 0.0) OR (fKpE < 0.0) THEN
    fTrimOut_pct := 0.0;        // 输出归 0 / Output zero
    bTensionAlarm := FALSE;     // 不误报超差 / No false alarm
    bEdgeAlarm := FALSE;        // 报警复位 / Alarm reset
    eErr := 16#0003_03D6;       // 故障码 / Fault code
    RETURN;                     // 本拍结束 / End of cycle
END_IF

// ---- 首扫初始化（R16 首扫纪律）/ First-scan initialization ----
IF xFirstScan THEN
    fTrimOut_pct := 0.0;        // 输出从 0 起步 / Output starts at zero
    xFirstScan := FALSE;        // 清标记 / Clear flag
END_IF

// ---- 权重钳位与归一（和恒为 1，不得双环各自满幅叠加）/ Weight clamp and normalize ----
fWeightTSafe := fWeightT;       // 原值 / As-is
IF fWeightTSafe < 0.0 THEN
    fWeightTSafe := 0.0;        // 下限 / Lower clamp
ELSIF fWeightTSafe > 1.0 THEN
    fWeightTSafe := 1.0;        // 上限 / Upper clamp
END_IF
fWeightE := 1.0 - fWeightTSafe; // 纠偏权重 / Edge weight

// ---- 容差兜底 / Tolerance fallbacks ----
IF fEdgeTol_mm <= 0.0 THEN
    fEdgeTolSafe := 0.1;        // 兜底 0.1 mm / Fallback 0.1 mm
ELSE
    fEdgeTolSafe := fEdgeTol_mm;    // 原值 / As-is
END_IF
IF fTensionTolPct <= 0.0 THEN
    fTolPctSafe := 0.5;         // 兜底 0.5 % / Fallback 0.5 %
ELSE
    fTolPctSafe := fTensionTolPct;  // 原值 / As-is
END_IF

// ---- 饱和故障锁存与解除 / Saturation latch and release ----
IF bSatLatch THEN
    fTrimOut_pct := 0.0;        // 锁存中输出归 0 / Zero output when latched
    bTensionAlarm := FALSE;     // 报警复位 / Alarm reset
    eErr := 16#0003_03D8;       // 故障码回放 / Fault code replay
    IF bReset THEN
        bSatLatch := FALSE;     // 解除锁存 / Release latch
    END_IF
    RETURN;                     // 本拍结束 / End of cycle
END_IF

// ---- 使能撤销：双环输出归 0 / Disable: outputs zero ----
IF NOT bEnable THEN
    fTrimOut_pct := 0.0;        // 输出归 0 / Output zero
    bTensionAlarm := FALSE;     // 报警复位 / Alarm reset
    bEdgeAlarm := FALSE;        // 报警复位 / Alarm reset
    eErr := 16#0003_03D4;       // 信息级：空闲 / Info: idle
    RETURN;                     // 本拍结束 / End of cycle
END_IF

// ---- 偏差计算 / Deviation computation ----
fDev_N := fTensionSp_N - fTension_N;        // 张力偏差 / Tension deviation [N]
fEdgeDev_mm := fEdgePos_mm - fEdgeCenter_mm;    // 边缘偏差 / Edge deviation [mm]

// ---- 张力超差报警（分母有设定值闸，sp>0 已由组态闸保证）/ Tension alarm ----
bTensionAlarm := (ABS(fDev_N) / fTensionSp_N * 100.0 > fTolPctSafe);   // 超差判 / Over-tolerance

// ---- 边缘跑偏报警 / Edge alarm ----
bEdgeAlarm := (ABS(fEdgeDev_mm) > fEdgeTolSafe);    // 跑偏判 / Over-tolerance

// ---- 网带停止：双环输出归 0，积分保持（再启动无扰）/ Web stopped: outputs zero, hold ----
IF NOT bWebRun THEN
    fTrimOut_pct := 0.0;        // 输出归 0 / Output zero
    eErr := 16#0003_03D7;       // 信息级：停机冻结 / Info: stopped freeze
    RETURN;                     // 本拍结束 / End of cycle
END_IF

// ---- 双环计算 / Dual loop computation ----
fTensionTrim := fWeightTSafe * fKpT * fDev_N;       // 张力项（跑偏报警时冻结）/ Tension term
fEdgeTrim := fWeightE * fKpE * fEdgeDev_mm;         // 纠偏项 / Edge term

IF bEdgeAlarm THEN
    // 跑偏超差：张力环输出冻结以免叠加扰动，输出只含纠偏项 / Edge alarm: tension frozen
    fTrimOut_pct := fEdgeTrim;  // 只含纠偏项 / Edge term only
    eErr := 16#0003_03D7;       // 信息级：张力环冻结 / Info: tension frozen
ELSE
    fTrimOut_pct := fTensionTrim + fEdgeTrim;   // 双环加权合成 / Weighted sum
    eErr := 16#0003_03D4;       // 信息级：双环正常 / Info: normal
END_IF

// ---- 输出限幅：先钳后使用 / Output clamp ----
IF fTrimOut_pct > fTrimMax_pct THEN
    fTrimOut_pct := fTrimMax_pct;   // 上限钳 / Upper clamp
ELSIF fTrimOut_pct < -fTrimMax_pct THEN
    fTrimOut_pct := -fTrimMax_pct;  // 下限钳 / Lower clamp
END_IF

// ---- 饱和监控：触限 + 同向偏差超容差 持续 10 s → 锁存 / Saturation monitor ----
bSatCond := FALSE;              // 条件复位 / Reset
IF (fTrimOut_pct >= fTrimMax_pct) AND (fDev_N > 0.0)
   AND (ABS(fDev_N) / fTensionSp_N * 100.0 > fTolPctSafe) THEN
    bSatCond := TRUE;           // 正向饱和 / Positive saturation
END_IF
IF (fTrimOut_pct <= -fTrimMax_pct) AND (fDev_N < 0.0)
   AND (ABS(fDev_N) / fTensionSp_N * 100.0 > fTolPctSafe) THEN
    bSatCond := TRUE;           // 负向饱和 / Negative saturation
END_IF
tonSat(IN := bSatCond, PT := T#10S);    // 定时器无条件周期刷新 / Unconditional refresh
IF tonSat.Q THEN
    bSatLatch := TRUE;          // 锁存 / Latch
    fTrimOut_pct := 0.0;        // 输出归 0 / Output zero
    eErr := 16#0003_03D8;       // 故障码 / Fault code
END_IF

END_FUNCTION_BLOCK

(* ---- FB_DL_GloveBoxAtmoCtrl.st ---- *)
(*
  FB_DL_GloveBoxAtmoCtrl  —  手套箱气氛联锁 / Glove-box atmosphere interlock control
  分类 Category : DL_Device
  码位 Code     : 16#03_2_06
  版本 Version  : 1.0.0
  溯源 Source   : NAMUR NE107 语义借鉴 · clean-room 实现，仅借分类/参数域/命名，未复制源码
  功能 Function : 1) 水/氧含量双路越限判定（带迟滞），任一路越限禁开门；
                  2) 开门许可经 FB_DL_InterlockMatrix 双条件联锁出口（复用）；
                  3) 净化循环请求与开门互斥仲裁；NE107 六态映射出口。
  边界 Boundary : ① 任一路无效按「越限」安全侧禁开门（R42 家族）；
                  ② 门限带迟滞防反复禁投；
                  ③ 越限解除须双路均回窗 + 最短维持时间（FB33-2 可达）；
                  ④ 净化请求与开门互斥仲裁（净化优先）；
                  ⑤ 未知状态归 eUnknown 绝不归 eOk；
                  ⑥ 输出三行同向：开门许可 → 净化请求 → NE107 态。
  依赖 Depends  : FB_DL_InterlockMatrix × 1（双条件联锁出口，每拍无条件调用）
                  E_DL_Ne107Status（属主件 I_DL_DeviceHealth，只引用不重声明）

  码表 Error codes（本件子码步进 16#10，避让邻件码位）:
    16#0002_0306 故障级：组态非法（门限倒置 / 迟滞 <= 0 / 维持时间 <= 0）
    16#0002_0316 故障级：相 ID 越界（枚举兜底路径）
    16#0002_0326 信息级：双路越限开门闭锁维持中 / 无效通道按越限处理（不置 bError）
*)

TYPE E_DL_GbaPhase :
(
    eIdle   := 0,  // 空闲 / Idle
    eWatch  := 10, // 气氛监视 / Atmosphere watching
    ePurge  := 20, // 净化循环请求保持 / Purge request held
    eFault  := 90  // 组态故障锁定 / Configuration fault locked
);
END_TYPE

FUNCTION_BLOCK FB_DL_GloveBoxAtmoCtrl
VAR_INPUT
    bEnable       : BOOL;                           // 总使能，FALSE 回空闲 / Master enable
    bReset        : BOOL;                           // 复位，上升沿清组态故障 / Reset, clears fault
    fH2oPpm       : REAL;                           // 水含量 [ppm] / Water content [ppm]
    fO2Ppm        : REAL;                           // 氧含量 [ppm] / Oxygen content [ppm]
    fH2oMaxPpm    : REAL := 5.0;                    // 水含量门限 [ppm] / Water limit [ppm]
    fO2MaxPpm     : REAL := 10.0;                   // 氧含量门限 [ppm] / Oxygen limit [ppm]
    fHystPpm      : REAL := 0.5;                    // 迟滞回差 [ppm]，域 > 0 / Hysteresis band [ppm]
    bDoorReq      : BOOL;                           // 开门请求 / Door request
    tSustainMin   : TIME := T#30S;                  // 回窗最短维持时间 [s]，域 > 0 / Min sustain time after back-in-window
    fEps          : REAL := 1.0E-6;                 // 浮点判零容差 [1] / Floating zero tolerance
END_VAR
VAR_OUTPUT
    bDoorPermit   : BOOL;                           // 开门许可出口（联锁矩阵放行）/ Door permit output
    bPurgeReq     : BOOL;                           // 净化循环请求（互斥仲裁后）/ Purge cycle request
    eNe107        : E_DL_Ne107Status;               // NE107 六态映射出口 / NE107 status mapping
    bError        : BOOL;                           // 故障标志，与故障级码配对 / Fault flag
    uErrorId      : UDINT;                          // 事件码，0 = 无事件 / Event code
    eStateOut     : E_DL_GbaPhase;                  // 状态机当前态，段尾单点映射 / Phase mapped at tail
END_VAR
VAR
    _eState       : E_DL_GbaPhase := E_DL_GbaPhase.eIdle;  // 内部状态 / Internal state
    fbIlk         : FB_DL_InterlockMatrix;          // 联锁矩阵实例（无条件调用）/ Interlock matrix instance
    rtrReset      : R_TRIG;                         // 复位沿 / Reset edge
    tonSustain    : TON;                            // 回窗维持计时器 / Back-in-window sustain timer
    abCondOk      : ARRAY[0..15] OF BOOL;           // 联锁条件表（ch0 水 / ch1 氧）/ Interlock condition table
    auInvertMask  : WORD;                           // 取反掩码（不取反）/ Invert mask
    auTripMask    : WORD;                           // 停机级掩码（双路均停机级）/ Trip-class mask
    bCfgOk        : BOOL;                           // 组态合法标志 / Configuration valid
    bH2oOk        : BOOL;                           // 水路本拍有效 / Water channel valid
    bO2Ok         : BOOL;                           // 氧路本拍有效 / Oxygen channel valid
    bH2oInWin     : BOOL;                           // 水路在窗（含迟滞）/ Water in window
    bO2InWin      : BOOL;                           // 氧路在窗（含迟滞）/ Oxygen in window
    bAnyOver      : BOOL;                           // 任一路越限或无效（电平）/ Any channel over or invalid
    bAllInWin     : BOOL;                           // 双路均在窗 / Both in window
    bSustainOk    : BOOL;                           // 维持时间已满足 / Sustain time met
    bHystWaterUp  : BOOL;                           // 水路迟滞越限状态（持有）/ Water over-limit hysteresis state
    bHystO2Up     : BOOL;                           // 氧路迟滞越限状态（持有）/ Oxygen over-limit hysteresis state
    uFault        : UDINT;                          // 锁存故障码 / Latched fault code
    uInfo         : UDINT;                          // 信息级码 / Information code
END_VAR
VAR CONSTANT
    DL_GBA_INFMAX : REAL := 1.0E30;                 // 含量有限值幅值上限 [ppm] / Content finite bound [ppm]
END_VAR

(* === 段 0 · 实例刷新 === *)
rtrReset(CLK := bReset);                          // 每拍刷新复位沿

(* === 段 1 · 组态闸 === *)
bCfgOk := (fH2oMaxPpm > fHystPpm) AND (fO2MaxPpm > fHystPpm)   // 门限须大于迟滞带（防带翻转）
          AND (fHystPpm > fEps)                   // 迟滞正域
          AND (TIME_TO_REAL(tSustainMin) > fEps)  // 维持时间正域
          AND (fH2oMaxPpm = fH2oMaxPpm) AND (fO2MaxPpm = fO2MaxPpm);  // NaN 自反
IF NOT bCfgOk THEN
    uFault := 16#0002_0306;                       // 故障级：组态非法
END_IF
IF rtrReset.Q AND bCfgOk THEN
    uFault := 16#0000;                            // 复位沿清锁存（解除路径可达）
END_IF
uInfo := 16#0000;                                 // 信息码每拍清零

(* === 段 2 · 双路域闸与迟滞越限判定 === *)
bH2oOk := (fH2oPpm = fH2oPpm) AND (fH2oPpm >= 0.0) AND (fH2oPpm < DL_GBA_INFMAX);  // 水路 NaN 自反 + 非负域
bO2Ok := (fO2Ppm = fO2Ppm) AND (fO2Ppm >= 0.0) AND (fO2Ppm < DL_GBA_INFMAX);       // 氧路域闸
IF bH2oOk THEN
    IF fH2oPpm >= fH2oMaxPpm THEN
        bHystWaterUp := TRUE;                     // 越门限置迟滞状态
    ELSIF fH2oPpm < fH2oMaxPpm - fHystPpm THEN
        bHystWaterUp := FALSE;                    // 回差带内解除（防反复禁投）
    END_IF
ELSE
    bHystWaterUp := TRUE;                         // 无效按越限安全侧（R42 家族）
    uInfo := 16#0002_0326;                        // 信息级：无效通道按越限处理
END_IF
IF bO2Ok THEN
    IF fO2Ppm >= fO2MaxPpm THEN
        bHystO2Up := TRUE;                        // 越门限置迟滞状态
    ELSIF fO2Ppm < fO2MaxPpm - fHystPpm THEN
        bHystO2Up := FALSE;                       // 回差带内解除
    END_IF
ELSE
    bHystO2Up := TRUE;                            // 无效按越限安全侧
    uInfo := 16#0002_0326;                        // 信息级：无效通道按越限处理
END_IF
bAnyOver := bHystWaterUp OR bHystO2Up;            // 任一路越限或无效
bAllInWin := (NOT bHystWaterUp) AND (NOT bHystO2Up);   // 双路均在窗

(* === 段 3 · 回窗最短维持时间（FB33-2：越限解除须回窗 + 最短维持）=== *)
tonSustain(IN := bAllInWin, PT := tSustainMin);   // 双路回窗才开始计时（越限即断输入复位）
bSustainOk := tonSustain.Q;                       // 维持时间满足
IF bAnyOver AND (NOT bAllInWin) THEN
    uInfo := 16#0002_0326;                        // 信息级：越限闭锁维持中
END_IF

(* === 段 4 · 联锁矩阵实例（无条件调用，双条件停机级）=== *)
abCondOk[0] := bH2oOk AND (NOT bHystWaterUp);     // 条件 0 = 水路有效且在窗
abCondOk[1] := bO2Ok AND (NOT bHystO2Up);         // 条件 1 = 氧路有效且在窗
auInvertMask := 16#0000;                          // 不取反
auTripMask := 16#0003;                            // 双路均停机级（bit0/bit1）
fbIlk(abConditionOk := abCondOk,                  // 条件表
      auInvertMask := auInvertMask,               // 取反掩码
      auTripMask := auTripMask,                   // 停机级掩码
      bEnable := bEnable AND bCfgOk,              // 使能透传
      bReset := rtrReset.Q);                      // 复位沿透传

(* === 段 5 · 主状态机（ENUM + CASE，含 ELSE 兜底）=== *)
CASE _eState OF
E_DL_GbaPhase.eIdle :
    IF uFault <> 16#0000 THEN
        _eState := E_DL_GbaPhase.eFault;          // 故障优先
    ELSIF bEnable AND bCfgOk AND bAnyOver THEN
        _eState := E_DL_GbaPhase.ePurge;          // 越限进净化请求相
    ELSIF bEnable AND bCfgOk THEN
        _eState := E_DL_GbaPhase.eWatch;          // 进监视相
    END_IF

E_DL_GbaPhase.eWatch :
    IF uFault <> 16#0000 THEN
        _eState := E_DL_GbaPhase.eFault;          // 故障转出
    ELSIF bAnyOver THEN
        _eState := E_DL_GbaPhase.ePurge;          // 越限转净化相
    END_IF

E_DL_GbaPhase.ePurge :
    IF uFault <> 16#0000 THEN
        _eState := E_DL_GbaPhase.eFault;          // 故障转出
    ELSIF bSustainOk AND (NOT bAnyOver) THEN
        _eState := E_DL_GbaPhase.eWatch;          // 双路回窗 + 维持满足：解除（路径可达）
    END_IF

E_DL_GbaPhase.eFault :
    IF uFault = 16#0000 THEN
        _eState := E_DL_GbaPhase.eIdle;           // 解锁回空闲
    END_IF

ELSE
    _eState := E_DL_GbaPhase.eFault;              // 非法状态拦截
    uFault := 16#0002_0316;                       // 故障级：相 ID 越界
END_CASE

(* === 段 6 · 输出映射（净化优先互斥仲裁）=== *)
bPurgeReq := (_eState = E_DL_GbaPhase.ePurge);    // 净化请求（净化相保持）
bDoorPermit := fbIlk.bPermitToRun AND bSustainOk AND (NOT bPurgeReq);   // 许可 = 矩阵放行 + 维持满足 + 与净化互斥
IF (NOT bH2oOk) OR (NOT bO2Ok) THEN
    eNe107 := E_DL_Ne107Status.eFailure;          // 任一路无效：失效态（信号不可信）
ELSIF bAnyOver THEN
    eNe107 := E_DL_Ne107Status.eOutOfSpec;        // 越限：超出规格态
ELSIF bPurgeReq THEN
    eNe107 := E_DL_Ne107Status.eCheckFunction;    // 净化循环中：功能检查态
ELSIF bEnable AND bCfgOk THEN
    eNe107 := E_DL_Ne107Status.eOk;               // 正常态
ELSE
    eNe107 := E_DL_Ne107Status.eUnknown;          // 未取得有效数据：未知态（绝不归 eOk）
END_IF
bError := (uFault <> 16#0000);                    // 故障标志仅由故障级码置位（R45 配对）
IF bError THEN
    uErrorId := uFault;                           // 故障级优先上报
ELSE
    uErrorId := uInfo;                            // 否则上报信息级码
END_IF
eStateOut := _eState;                             // 输出枚举段尾单点映射（N2 规则）
END_FUNCTION_BLOCK
